(* CODESYS project Example9_PLC.project

Project tree, tasks and I/O mapping:
  Device : CODESYS Control Win V3, 3S - Smart Software Solutions GmbH, order no. 305021, version 3.5.7.0
    application Application
      libraries: Standard, * (System)
      task MainTask (cyclic, interval t#20ms, priority 1) calls PLC_PRG
      program PLC_PRG [ST]
      global variables GVL
      function block FB_G4LTL [ST]
    Ethernet : Ethernet, 3S - Smart Software Solutions GmbH, version 3.5.7.0
      Modbus_TCP_Master : Modbus TCP Master, 3S - Smart Software Solutions GmbH, version 3.5.6.0
          settings: AutoReconnect = TRUE
        Modbus_TCP_Slave : Modbus TCP Slave, 3S - Smart Software Solutions GmbH, version 3.5.7.0
            settings: Unit-ID = 1; IPAddress = [127, 0, 0, 1]; Channel 0.Function Code = 4; Channel 0.Read Offset = 16#0000; Channel 0.Read Length = 1; Channel 0.Write Offset = 0; Channel 0.Write Length = 0; Channel 0.Cycle Time = 100; Channel 1.Function Code = 4; Channel 1.Read Offset = 16#0001; Channel 1.Read Length = 1; Channel 1.Write Offset = 0; Channel 1.Write Length = 0; Channel 1.Cycle Time = 100; Channel 2.Function Code = 4; Channel 2.Read Offset = 16#0002; Channel 2.Read Length = 1; Channel 2.Write Offset = 0; Channel 2.Write Length = 0; Channel 2.Cycle Time = 100; Channel 3.Function Code = 4; Channel 3.Read Offset = 16#0003; Channel 3.Read Length = 1; Channel 3.Write Offset = 0; Channel 3.Write Length = 0; Channel 3.Cycle Time = 100; Channel 4.Function Code = 4; Channel 4.Read Offset = 16#0004; Channel 4.Read Length = 1; Channel 4.Write Offset = 0; Channel 4.Write Length = 0; Channel 4.Cycle Time = 100; Channel 5.Function Code = 6; Channel 5.Read Offset = 0; Channel 5.Read Length = 0; Channel 5.Write Offset = 16#0000; Channel 5.Write Length = 1; Channel 5.Cycle Time = 100; Channel 6.Function Code = 6; Channel 6.Read Offset = 0;
              Channel 6.Read Length = 0; Channel 6.Write Offset = 16#0002; Channel 6.Write Length = 1; Channel 6.Cycle Time = 100; Channel 7.Function Code = 6; Channel 7.Read Offset = 0; Channel 7.Read Length = 0; Channel 7.Write Offset = 16#0003; Channel 7.Write Length = 1; Channel 7.Cycle Time = 100; Channel 8.Function Code = 6; Channel 8.Read Offset = 0; Channel 8.Read Length = 0; Channel 8.Write Offset = 16#0004; Channel 8.Write Length = 1; Channel 8.Cycle Time = 100; Channel 9.Function Code = 6; Channel 9.Read Offset = 0; Channel 9.Read Length = 0; Channel 9.Write Offset = 16#0001; Channel 9.Write Length = 1; Channel 9.Cycle Time = 100
            input  Application.dIn0 : BOOL  // Channel 0.Channel 0.Bit0
            input  Application.dIn1 : BOOL  // Channel 1.Channel 1.Bit0
            input  Application.dIn2 : BOOL  // Channel 2.Channel 2.Bit0
            input  Application.dIn3 : BOOL  // Channel 3.Channel 3.Bit0
            input  Application.dIn4 : BOOL  // Channel 4.Channel 4.Bit0
            output Application.dOut0 : BOOL  // Channel 5.Channel 5.Bit0
            output Application.dOut2 : BOOL  // Channel 6.Channel 6.Bit0
            output Application.dOut3 : BOOL  // Channel 7.Channel 7.Bit0
            output Application.dOut4 : BOOL  // Channel 8.Channel 8.Bit0
            output Application.dOut1 : BOOL  // Channel 9.Channel 9.Bit0
            unmapped channels: Channel 0, Channel 1, Channel 2, Channel 3, Channel 4, Channel 5, Channel 6, Channel 7, Channel 8, Channel 9
*)

// Device/Application/GVL
VAR_GLOBAL
	
dIn0 : BOOL;
dIn1 : BOOL;
dIn2 : BOOL;
dIn3 : BOOL;
dIn4 : BOOL;

dOut0 : BOOL;
dOut1 : BOOL; 
dOut2 : BOOL; 
dOut3 : BOOL; 
dOut4 : BOOL; 
END_VAR

// Device/Application/PLC_PRG
PROGRAM PLC_PRG
VAR 
	fb: FB_G4LTL;	
END_VAR



// Direct looping
// Assign pins (from global variable to function block) 
fb.x0 := dIn0;

// Assign pins (from function block to global variable)
dOut0 := fb.y0;
dOut1 := fb.y1;
dOut2 := fb.y2;

// Run the function block
fb();

END_PROGRAM

// Device/Application/FB_G4LTL
FUNCTION_BLOCK FB_G4LTL
 (* Variable definition *)
   VAR_INPUT
      x0	: BOOL;
   END_VAR
   VAR_OUTPUT
      y0	: BOOL;
      y1	: BOOL;
      y2	: BOOL;
   END_VAR
   VAR
   (* The total number of states equals to 11 *)
      cstate16	: LINT := 0;
      t0	: TON;
      t0_reset	: BOOL := FALSE;
      t0_up	: BOOL := FALSE;
      t0_start	: BOOL := FALSE;
      t1	: TON;
      t1_reset	: BOOL := FALSE;
      t1_up	: BOOL := FALSE;
      t1_start	: BOOL := FALSE;	  
	  
	  T0_VALUE	: TIME := TIME#10S;
      T1_VALUE	: TIME := TIME#5s;
   END_VAR
   (* Constant definition  *)

CASE cstate16 OF
48641:
    IF ((x0 = FALSE) AND  (t0.Q = FALSE) AND  (t1.Q = FALSE)) THEN 
        cstate16 := 34931; y0 := FALSE; y1 := FALSE; y2 := FALSE; t0_start := FALSE;t1_start := FALSE; 
    ELSIF ((x0 = FALSE) AND  (t0.Q = FALSE) AND  (t1.Q = TRUE)) THEN 
        cstate16 := 34932; y0 := FALSE; y1 := FALSE; y2 := FALSE; t0_start := FALSE;t1_start := FALSE; 
    ELSIF ((x0 = FALSE) AND  (t0.Q = TRUE) AND  (t1.Q = FALSE)) THEN 
        cstate16 := 27731; y0 := FALSE; y1 := FALSE; y2 := FALSE; t0_start := FALSE;t1_start := TRUE; t1_up := FALSE; 
    ELSIF ((x0 = FALSE) AND  (t0.Q = TRUE) AND  (t1.Q = TRUE)) THEN 
        cstate16 := 27732; y0 := FALSE; y1 := FALSE; y2 := FALSE; t0_start := FALSE;t1_start := TRUE; t1_up := FALSE; 
    ELSIF ((x0 = TRUE) AND  (t0.Q = FALSE) AND  (t1.Q = FALSE)) THEN 
        cstate16 := 48641; y0 := TRUE; y1 := TRUE; y2 := FALSE; t0_start := FALSE;t1_start := FALSE; 
    ELSIF ((x0 = TRUE) AND  (t0.Q = FALSE) AND  (t1.Q = TRUE)) THEN 
        cstate16 := 48646; y0 := TRUE; y1 := TRUE; y2 := TRUE; t0_start := FALSE;t1_start := FALSE; 
    ELSIF ((x0 = TRUE) AND  (t0.Q = TRUE) AND  (t1.Q = FALSE)) THEN 
        cstate16 := 42449; y0 := TRUE; y1 := TRUE; y2 := FALSE; t0_start := FALSE;t1_start := TRUE; t1_up := FALSE; 
    ELSIF ((x0 = TRUE) AND  (t0.Q = TRUE) AND  (t1.Q = TRUE)) THEN 
        cstate16 := 42453; y0 := TRUE; y1 := TRUE; y2 := TRUE; t0_start := FALSE;t1_start := TRUE; t1_up := FALSE; 
    END_IF;
46659:
    IF ((x0 = FALSE) AND  (t0.Q = FALSE) AND  (t1.Q = FALSE)) THEN 
        cstate16 := 32883; y0 := FALSE; y1 := FALSE; y2 := FALSE; t0_start := FALSE;t1_start := FALSE; 
    ELSIF ((x0 = FALSE) AND  (t0.Q = FALSE) AND  (t1.Q = TRUE)) THEN 
        cstate16 := 34932; y0 := FALSE; y1 := FALSE; y2 := FALSE; t0_start := FALSE;t1_start := FALSE; 
    ELSIF ((x0 = FALSE) AND  (t0.Q = TRUE) AND  (t1.Q = FALSE)) THEN 
        cstate16 := 27763; y0 := FALSE; y1 := FALSE; y2 := FALSE; t0_start := FALSE;t1_start := FALSE; 
    ELSIF ((x0 = FALSE) AND  (t0.Q = TRUE) AND  (t1.Q = TRUE)) THEN 
        cstate16 := 28788; y0 := FALSE; y1 := FALSE; y2 := FALSE; t0_start := FALSE;t1_start := FALSE; 
    ELSIF ((x0 = TRUE) AND  (t0.Q = FALSE) AND  (t1.Q = FALSE)) THEN 
        cstate16 := 41187; y0 := TRUE; y1 := FALSE; y2 := FALSE; t0_start := TRUE; t0_up := FALSE;t1_start := FALSE; 
    ELSIF ((x0 = TRUE) AND  (t0.Q = FALSE) AND  (t1.Q = TRUE)) THEN 
        cstate16 := 40167; y0 := TRUE; y1 := FALSE; y2 := TRUE; t0_start := TRUE; t0_up := FALSE;t1_start := FALSE; 
    ELSIF ((x0 = TRUE) AND  (t0.Q = TRUE) AND  (t1.Q = FALSE)) THEN 
        cstate16 := 46659; y0 := TRUE; y1 := FALSE; y2 := FALSE; t0_start := FALSE;t1_start := FALSE; 
    ELSIF ((x0 = TRUE) AND  (t0.Q = TRUE) AND  (t1.Q = TRUE)) THEN 
        cstate16 := 47687; y0 := TRUE; y1 := FALSE; y2 := TRUE; t0_start := FALSE;t1_start := FALSE; 
    END_IF;
46651:
    IF ((x0 = FALSE) AND  (t0.Q = FALSE) AND  (t1.Q = FALSE)) THEN 
        cstate16 := 32883; y0 := FALSE; y1 := FALSE; y2 := FALSE; t0_start := FALSE;t1_start := FALSE; 
    ELSIF ((x0 = FALSE) AND  (t0.Q = FALSE) AND  (t1.Q = TRUE)) THEN 
        cstate16 := 34932; y0 := FALSE; y1 := FALSE; y2 := FALSE; t0_start := FALSE;t1_start := FALSE; 
    ELSIF ((x0 = FALSE) AND  (t0.Q = TRUE) AND  (t1.Q = FALSE)) THEN 
        cstate16 := 27763; y0 := FALSE; y1 := FALSE; y2 := FALSE; t0_start := FALSE;t1_start := FALSE; 
    ELSIF ((x0 = FALSE) AND  (t0.Q = TRUE) AND  (t1.Q = TRUE)) THEN 
        cstate16 := 28788; y0 := FALSE; y1 := FALSE; y2 := FALSE; t0_start := FALSE;t1_start := FALSE; 
    ELSIF ((x0 = TRUE) AND  (t0.Q = FALSE) AND  (t1.Q = FALSE)) THEN 
        cstate16 := 41643; y0 := TRUE; y1 := TRUE; y2 := TRUE; t0_start := TRUE; t0_up := FALSE;t1_start := FALSE; 
    ELSIF ((x0 = TRUE) AND  (t0.Q = FALSE) AND  (t1.Q = TRUE)) THEN 
        cstate16 := 40647; y0 := TRUE; y1 := TRUE; y2 := TRUE; t0_start := TRUE; t0_up := FALSE;t1_start := FALSE; 
    ELSIF ((x0 = TRUE) AND  (t0.Q = TRUE) AND  (t1.Q = FALSE)) THEN 
        cstate16 := 46747; y0 := TRUE; y1 := TRUE; y2 := TRUE; t0_start := FALSE;t1_start := FALSE; 
    ELSIF ((x0 = TRUE) AND  (t0.Q = TRUE) AND  (t1.Q = TRUE)) THEN 
        cstate16 := 47799; y0 := TRUE; y1 := TRUE; y2 := TRUE; t0_start := FALSE;t1_start := FALSE; 
    END_IF;
25798:
    IF ((x0 = FALSE) AND  (t0.Q = FALSE) AND  (t1.Q = FALSE)) THEN 
        cstate16 := 26739; y0 := FALSE; y1 := FALSE; y2 := FALSE; t0_start := FALSE;t1_start := FALSE; 
    ELSIF ((x0 = FALSE) AND  (t0.Q = FALSE) AND  (t1.Q = TRUE)) THEN 
        cstate16 := 26740; y0 := FALSE; y1 := FALSE; y2 := FALSE; t0_start := FALSE;t1_start := FALSE; 
    ELSIF ((x0 = FALSE) AND  (t0.Q = TRUE) AND  (t1.Q = FALSE)) THEN 
        cstate16 := 17491; y0 := FALSE; y1 := FALSE; y2 := FALSE; t0_start := FALSE;t1_start := TRUE; t1_up := FALSE; 
    ELSIF ((x0 = FALSE) AND  (t0.Q = TRUE) AND  (t1.Q = TRUE)) THEN 
        cstate16 := 17492; y0 := FALSE; y1 := FALSE; y2 := FALSE; t0_start := FALSE;t1_start := TRUE; t1_up := FALSE; 
    ELSIF ((x0 = TRUE) AND  (t0.Q = FALSE) AND  (t1.Q = FALSE)) THEN 
        cstate16 := 26042; y0 := TRUE; y1 := FALSE; y2 := TRUE; t0_start := FALSE;t1_start := FALSE; 
    ELSIF ((x0 = TRUE) AND  (t0.Q = FALSE) AND  (t1.Q = TRUE)) THEN 
        cstate16 := 26038; y0 := TRUE; y1 := FALSE; y2 := TRUE; t0_start := FALSE;t1_start := FALSE; 
    ELSIF ((x0 = TRUE) AND  (t0.Q = TRUE) AND  (t1.Q = FALSE)) THEN 
        cstate16 := 42457; y0 := TRUE; y1 := TRUE; y2 := TRUE; t0_start := FALSE;t1_start := TRUE; t1_up := FALSE; 
    ELSIF ((x0 = TRUE) AND  (t0.Q = TRUE) AND  (t1.Q = TRUE)) THEN 
        cstate16 := 42453; y0 := TRUE; y1 := TRUE; y2 := TRUE; t0_start := FALSE;t1_start := TRUE; t1_up := FALSE; 
    END_IF;
34931:
    IF ((x0 = FALSE) AND  (t0.Q = FALSE) AND  (t1.Q = FALSE)) THEN 
        cstate16 := 34931; y0 := FALSE; y1 := FALSE; y2 := FALSE; t0_start := FALSE;t1_start := FALSE; 
    ELSIF ((x0 = FALSE) AND  (t0.Q = FALSE) AND  (t1.Q = TRUE)) THEN 
        cstate16 := 34932; y0 := FALSE; y1 := FALSE; y2 := FALSE; t0_start := FALSE;t1_start := FALSE; 
    ELSIF ((x0 = FALSE) AND  (t0.Q = TRUE) AND  (t1.Q = FALSE)) THEN 
        cstate16 := 27731; y0 := FALSE; y1 := FALSE; y2 := FALSE; t0_start := FALSE;t1_start := TRUE; t1_up := FALSE; 
    ELSIF ((x0 = FALSE) AND  (t0.Q = TRUE) AND  (t1.Q = TRUE)) THEN 
        cstate16 := 27732; y0 := FALSE; y1 := FALSE; y2 := FALSE; t0_start := FALSE;t1_start := TRUE; t1_up := FALSE; 
    ELSIF ((x0 = TRUE) AND  (t0.Q = FALSE) AND  (t1.Q = FALSE)) THEN 
        cstate16 := 40163; y0 := TRUE; y1 := FALSE; y2 := FALSE; t0_start := TRUE; t0_up := FALSE;t1_start := FALSE; 
    ELSIF ((x0 = TRUE) AND  (t0.Q = FALSE) AND  (t1.Q = TRUE)) THEN 
        cstate16 := 40167; y0 := TRUE; y1 := FALSE; y2 := TRUE; t0_start := TRUE; t0_up := FALSE;t1_start := FALSE; 
    ELSIF ((x0 = TRUE) AND  (t0.Q = TRUE) AND  (t1.Q = FALSE)) THEN 
        cstate16 := 38147; y0 := TRUE; y1 := TRUE; y2 := FALSE; t0_start := TRUE; t0_up := FALSE;t1_start := TRUE; t1_up := FALSE; 
    ELSIF ((x0 = TRUE) AND  (t0.Q = TRUE) AND  (t1.Q = TRUE)) THEN 
        cstate16 := 38152; y0 := TRUE; y1 := TRUE; y2 := TRUE; t0_start := TRUE; t0_up := FALSE;t1_start := TRUE; t1_up := FALSE; 
    END_IF;
47687:
    IF ((x0 = FALSE) AND  (t0.Q = FALSE) AND  (t1.Q = FALSE)) THEN 
        cstate16 := 34931; y0 := FALSE; y1 := FALSE; y2 := FALSE; t0_start := FALSE;t1_start := FALSE; 
    ELSIF ((x0 = FALSE) AND  (t0.Q = FALSE) AND  (t1.Q = TRUE)) THEN 
        cstate16 := 34932; y0 := FALSE; y1 := FALSE; y2 := FALSE; t0_start := FALSE;t1_start := FALSE; 
    ELSIF ((x0 = FALSE) AND  (t0.Q = TRUE) AND  (t1.Q = FALSE)) THEN 
        cstate16 := 28787; y0 := FALSE; y1 := FALSE; y2 := FALSE; t0_start := FALSE;t1_start := FALSE; 
    ELSIF ((x0 = FALSE) AND  (t0.Q = TRUE) AND  (t1.Q = TRUE)) THEN 
        cstate16 := 28788; y0 := FALSE; y1 := FALSE; y2 := FALSE; t0_start := FALSE;t1_start := FALSE; 
    ELSIF ((x0 = TRUE) AND  (t0.Q = FALSE) AND  (t1.Q = FALSE)) THEN 
        cstate16 := 40172; y0 := TRUE; y1 := FALSE; y2 := TRUE; t0_start := TRUE; t0_up := FALSE;t1_start := FALSE; 
    ELSIF ((x0 = TRUE) AND  (t0.Q = FALSE) AND  (t1.Q = TRUE)) THEN 
        cstate16 := 40167; y0 := TRUE; y1 := FALSE; y2 := TRUE; t0_start := TRUE; t0_up := FALSE;t1_start := FALSE; 
    ELSIF ((x0 = TRUE) AND  (t0.Q = TRUE) AND  (t1.Q = FALSE)) THEN 
        cstate16 := 47692; y0 := TRUE; y1 := FALSE; y2 := TRUE; t0_start := FALSE;t1_start := FALSE; 
    ELSIF ((x0 = TRUE) AND  (t0.Q = TRUE) AND  (t1.Q = TRUE)) THEN 
        cstate16 := 47687; y0 := TRUE; y1 := FALSE; y2 := TRUE; t0_start := FALSE;t1_start := FALSE; 
    END_IF;
43409:
    IF ((x0 = FALSE) AND  (t0.Q = FALSE) AND  (t1.Q = FALSE)) THEN 
        cstate16 := 34931; y0 := FALSE; y1 := FALSE; y2 := FALSE; t0_start := FALSE;t1_start := FALSE; 
    ELSIF ((x0 = FALSE) AND  (t0.Q = FALSE) AND  (t1.Q = TRUE)) THEN 
        cstate16 := 34932; y0 := FALSE; y1 := FALSE; y2 := FALSE; t0_start := FALSE;t1_start := FALSE; 
    ELSIF ((x0 = FALSE) AND  (t0.Q = TRUE) AND  (t1.Q = FALSE)) THEN 
        cstate16 := 28787; y0 := FALSE; y1 := FALSE; y2 := FALSE; t0_start := FALSE;t1_start := FALSE; 
    ELSIF ((x0 = FALSE) AND  (t0.Q = TRUE) AND  (t1.Q = TRUE)) THEN 
        cstate16 := 28788; y0 := FALSE; y1 := FALSE; y2 := FALSE; t0_start := FALSE;t1_start := FALSE; 
    ELSIF ((x0 = TRUE) AND  (t0.Q = FALSE) AND  (t1.Q = FALSE)) THEN 
        cstate16 := 48529; y0 := TRUE; y1 := FALSE; y2 := FALSE; t0_start := FALSE;t1_start := FALSE; 
    ELSIF ((x0 = TRUE) AND  (t0.Q = FALSE) AND  (t1.Q = TRUE)) THEN 
        cstate16 := 48534; y0 := TRUE; y1 := FALSE; y2 := TRUE; t0_start := FALSE;t1_start := FALSE; 
    ELSIF ((x0 = TRUE) AND  (t0.Q = TRUE) AND  (t1.Q = FALSE)) THEN 
        cstate16 := 43409; y0 := TRUE; y1 := FALSE; y2 := FALSE; t0_start := FALSE;t1_start := FALSE; 
    ELSIF ((x0 = TRUE) AND  (t0.Q = TRUE) AND  (t1.Q = TRUE)) THEN 
        cstate16 := 43414; y0 := TRUE; y1 := FALSE; y2 := TRUE; t0_start := FALSE;t1_start := FALSE; 
    END_IF;
34932:
    IF ((x0 = FALSE) AND  (t0.Q = FALSE) AND  (t1.Q = FALSE)) THEN 
        cstate16 := 34931; y0 := FALSE; y1 := FALSE; y2 := FALSE; t0_start := FALSE;t1_start := FALSE; 
    ELSIF ((x0 = FALSE) AND  (t0.Q = FALSE) AND  (t1.Q = TRUE)) THEN 
        cstate16 := 34932; y0 := FALSE; y1 := FALSE; y2 := FALSE; t0_start := FALSE;t1_start := FALSE; 
    ELSIF ((x0 = FALSE) AND  (t0.Q = TRUE) AND  (t1.Q = FALSE)) THEN 
        cstate16 := 27731; y0 := FALSE; y1 := FALSE; y2 := FALSE; t0_start := FALSE;t1_start := TRUE; t1_up := FALSE; 
    ELSIF ((x0 = FALSE) AND  (t0.Q = TRUE) AND  (t1.Q = TRUE)) THEN 
        cstate16 := 27732; y0 := FALSE; y1 := FALSE; y2 := FALSE; t0_start := FALSE;t1_start := TRUE; t1_up := FALSE; 
    ELSIF ((x0 = TRUE) AND  (t0.Q = FALSE) AND  (t1.Q = FALSE)) THEN 
        cstate16 := 40163; y0 := TRUE; y1 := FALSE; y2 := FALSE; t0_start := TRUE; t0_up := FALSE;t1_start := FALSE; 
    ELSIF ((x0 = TRUE) AND  (t0.Q = FALSE) AND  (t1.Q = TRUE)) THEN 
        cstate16 := 40164; y0 := TRUE; y1 := FALSE; y2 := FALSE; t0_start := TRUE; t0_up := FALSE;t1_start := FALSE; 
    ELSIF ((x0 = TRUE) AND  (t0.Q = TRUE) AND  (t1.Q = FALSE)) THEN 
        cstate16 := 38147; y0 := TRUE; y1 := TRUE; y2 := FALSE; t0_start := TRUE; t0_up := FALSE;t1_start := TRUE; t1_up := FALSE; 
    ELSIF ((x0 = TRUE) AND  (t0.Q = TRUE) AND  (t1.Q = TRUE)) THEN 
        cstate16 := 38148; y0 := TRUE; y1 := TRUE; y2 := FALSE; t0_start := TRUE; t0_up := FALSE;t1_start := TRUE; t1_up := FALSE; 
    END_IF;
6209:
    IF ((x0 = FALSE) AND  (t0.Q = FALSE) AND  (t1.Q = FALSE)) THEN 
        cstate16 := 34931; y0 := FALSE; y1 := FALSE; y2 := FALSE; t0_start := FALSE;t1_start := FALSE; 
    ELSIF ((x0 = FALSE) AND  (t0.Q = FALSE) AND  (t1.Q = TRUE)) THEN 
        cstate16 := 34932; y0 := FALSE; y1 := FALSE; y2 := FALSE; t0_start := FALSE;t1_start := FALSE; 
    ELSIF ((x0 = FALSE) AND  (t0.Q = TRUE) AND  (t1.Q = FALSE)) THEN 
        cstate16 := 28787; y0 := FALSE; y1 := FALSE; y2 := FALSE; t0_start := FALSE;t1_start := FALSE; 
    ELSIF ((x0 = FALSE) AND  (t0.Q = TRUE) AND  (t1.Q = TRUE)) THEN 
        cstate16 := 28788; y0 := FALSE; y1 := FALSE; y2 := FALSE; t0_start := FALSE;t1_start := FALSE; 
    ELSIF ((x0 = TRUE) AND  (t0.Q = FALSE) AND  (t1.Q = FALSE)) THEN 
        cstate16 := 14401; y0 := FALSE; y1 := FALSE; y2 := FALSE; t0_start := FALSE;t1_start := FALSE; 
    ELSIF ((x0 = TRUE) AND  (t0.Q = FALSE) AND  (t1.Q = TRUE)) THEN 
        cstate16 := 14406; y0 := FALSE; y1 := FALSE; y2 := TRUE; t0_start := FALSE;t1_start := FALSE; 
    ELSIF ((x0 = TRUE) AND  (t0.Q = TRUE) AND  (t1.Q = FALSE)) THEN 
        cstate16 := 6209; y0 := FALSE; y1 := FALSE; y2 := FALSE; t0_start := FALSE;t1_start := FALSE; 
    ELSIF ((x0 = TRUE) AND  (t0.Q = TRUE) AND  (t1.Q = TRUE)) THEN 
        cstate16 := 6214; y0 := FALSE; y1 := FALSE; y2 := TRUE; t0_start := FALSE;t1_start := FALSE; 
    END_IF;
42489:
    IF ((x0 = FALSE) AND  (t0.Q = FALSE) AND  (t1.Q = FALSE)) THEN 
        cstate16 := 32883; y0 := FALSE; y1 := FALSE; y2 := FALSE; t0_start := FALSE;t1_start := FALSE; 
    ELSIF ((x0 = FALSE) AND  (t0.Q = FALSE) AND  (t1.Q = TRUE)) THEN 
        cstate16 := 34932; y0 := FALSE; y1 := FALSE; y2 := FALSE; t0_start := FALSE;t1_start := FALSE; 
    ELSIF ((x0 = FALSE) AND  (t0.Q = TRUE) AND  (t1.Q = FALSE)) THEN 
        cstate16 := 27763; y0 := FALSE; y1 := FALSE; y2 := FALSE; t0_start := FALSE;t1_start := FALSE; 
    ELSIF ((x0 = FALSE) AND  (t0.Q = TRUE) AND  (t1.Q = TRUE)) THEN 
        cstate16 := 28788; y0 := FALSE; y1 := FALSE; y2 := FALSE; t0_start := FALSE;t1_start := FALSE; 
    ELSIF ((x0 = TRUE) AND  (t0.Q = FALSE) AND  (t1.Q = FALSE)) THEN 
        cstate16 := 49657; y0 := TRUE; y1 := TRUE; y2 := TRUE; t0_start := FALSE;t1_start := FALSE; 
    ELSIF ((x0 = TRUE) AND  (t0.Q = FALSE) AND  (t1.Q = TRUE)) THEN 
        cstate16 := 48646; y0 := TRUE; y1 := TRUE; y2 := TRUE; t0_start := FALSE;t1_start := FALSE; 
    ELSIF ((x0 = TRUE) AND  (t0.Q = TRUE) AND  (t1.Q = FALSE)) THEN 
        cstate16 := 42489; y0 := TRUE; y1 := TRUE; y2 := TRUE; t0_start := FALSE;t1_start := FALSE; 
    ELSIF ((x0 = TRUE) AND  (t0.Q = TRUE) AND  (t1.Q = TRUE)) THEN 
        cstate16 := 43526; y0 := TRUE; y1 := TRUE; y2 := TRUE; t0_start := FALSE;t1_start := FALSE; 
    END_IF;
6490:
    IF ((x0 = FALSE) AND  (t0.Q = FALSE) AND  (t1.Q = FALSE)) THEN 
        cstate16 := 34931; y0 := FALSE; y1 := FALSE; y2 := FALSE; t0_start := FALSE;t1_start := FALSE; 
    ELSIF ((x0 = FALSE) AND  (t0.Q = FALSE) AND  (t1.Q = TRUE)) THEN 
        cstate16 := 34932; y0 := FALSE; y1 := FALSE; y2 := FALSE; t0_start := FALSE;t1_start := FALSE; 
    ELSIF ((x0 = FALSE) AND  (t0.Q = TRUE) AND  (t1.Q = FALSE)) THEN 
        cstate16 := 28787; y0 := FALSE; y1 := FALSE; y2 := FALSE; t0_start := FALSE;t1_start := FALSE; 
    ELSIF ((x0 = FALSE) AND  (t0.Q = TRUE) AND  (t1.Q = TRUE)) THEN 
        cstate16 := 28788; y0 := FALSE; y1 := FALSE; y2 := FALSE; t0_start := FALSE;t1_start := FALSE; 
    ELSIF ((x0 = TRUE) AND  (t0.Q = FALSE) AND  (t1.Q = FALSE)) THEN 
        cstate16 := 14682; y0 := FALSE; y1 := TRUE; y2 := TRUE; t0_start := FALSE;t1_start := FALSE; 
    ELSIF ((x0 = TRUE) AND  (t0.Q = FALSE) AND  (t1.Q = TRUE)) THEN 
        cstate16 := 14678; y0 := FALSE; y1 := TRUE; y2 := TRUE; t0_start := FALSE;t1_start := FALSE; 
    ELSIF ((x0 = TRUE) AND  (t0.Q = TRUE) AND  (t1.Q = FALSE)) THEN 
        cstate16 := 6490; y0 := FALSE; y1 := TRUE; y2 := TRUE; t0_start := FALSE;t1_start := FALSE; 
    ELSIF ((x0 = TRUE) AND  (t0.Q = TRUE) AND  (t1.Q = TRUE)) THEN 
        cstate16 := 6486; y0 := FALSE; y1 := TRUE; y2 := TRUE; t0_start := FALSE;t1_start := FALSE; 
    END_IF;
6210:
    IF ((x0 = FALSE) AND  (t0.Q = FALSE) AND  (t1.Q = FALSE)) THEN 
        cstate16 := 34931; y0 := FALSE; y1 := FALSE; y2 := FALSE; t0_start := FALSE;t1_start := FALSE; 
    ELSIF ((x0 = FALSE) AND  (t0.Q = FALSE) AND  (t1.Q = TRUE)) THEN 
        cstate16 := 34932; y0 := FALSE; y1 := FALSE; y2 := FALSE; t0_start := FALSE;t1_start := FALSE; 
    ELSIF ((x0 = FALSE) AND  (t0.Q = TRUE) AND  (t1.Q = FALSE)) THEN 
        cstate16 := 28787; y0 := FALSE; y1 := FALSE; y2 := FALSE; t0_start := FALSE;t1_start := FALSE; 
    ELSIF ((x0 = FALSE) AND  (t0.Q = TRUE) AND  (t1.Q = TRUE)) THEN 
        cstate16 := 28788; y0 := FALSE; y1 := FALSE; y2 := FALSE; t0_start := FALSE;t1_start := FALSE; 
    ELSIF ((x0 = TRUE) AND  (t0.Q = FALSE) AND  (t1.Q = FALSE)) THEN 
        cstate16 := 14401; y0 := FALSE; y1 := FALSE; y2 := FALSE; t0_start := FALSE;t1_start := FALSE; 
    ELSIF ((x0 = TRUE) AND  (t0.Q = FALSE) AND  (t1.Q = TRUE)) THEN 
        cstate16 := 14402; y0 := FALSE; y1 := FALSE; y2 := FALSE; t0_start := FALSE;t1_start := FALSE; 
    ELSIF ((x0 = TRUE) AND  (t0.Q = TRUE) AND  (t1.Q = FALSE)) THEN 
        cstate16 := 6209; y0 := FALSE; y1 := FALSE; y2 := FALSE; t0_start := FALSE;t1_start := FALSE; 
    ELSIF ((x0 = TRUE) AND  (t0.Q = TRUE) AND  (t1.Q = TRUE)) THEN 
        cstate16 := 6210; y0 := FALSE; y1 := FALSE; y2 := FALSE; t0_start := FALSE;t1_start := FALSE; 
    END_IF;
25794:
    IF ((x0 = FALSE) AND  (t0.Q = FALSE) AND  (t1.Q = FALSE)) THEN 
        cstate16 := 26739; y0 := FALSE; y1 := FALSE; y2 := FALSE; t0_start := FALSE;t1_start := FALSE; 
    ELSIF ((x0 = FALSE) AND  (t0.Q = FALSE) AND  (t1.Q = TRUE)) THEN 
        cstate16 := 26740; y0 := FALSE; y1 := FALSE; y2 := FALSE; t0_start := FALSE;t1_start := FALSE; 
    ELSIF ((x0 = FALSE) AND  (t0.Q = TRUE) AND  (t1.Q = FALSE)) THEN 
        cstate16 := 17491; y0 := FALSE; y1 := FALSE; y2 := FALSE; t0_start := FALSE;t1_start := TRUE; t1_up := FALSE; 
    ELSIF ((x0 = FALSE) AND  (t0.Q = TRUE) AND  (t1.Q = TRUE)) THEN 
        cstate16 := 17492; y0 := FALSE; y1 := FALSE; y2 := FALSE; t0_start := FALSE;t1_start := TRUE; t1_up := FALSE; 
    ELSIF ((x0 = TRUE) AND  (t0.Q = FALSE) AND  (t1.Q = FALSE)) THEN 
        cstate16 := 26033; y0 := TRUE; y1 := FALSE; y2 := FALSE; t0_start := FALSE;t1_start := FALSE; 
    ELSIF ((x0 = TRUE) AND  (t0.Q = FALSE) AND  (t1.Q = TRUE)) THEN 
        cstate16 := 26034; y0 := TRUE; y1 := FALSE; y2 := FALSE; t0_start := FALSE;t1_start := FALSE; 
    ELSIF ((x0 = TRUE) AND  (t0.Q = TRUE) AND  (t1.Q = FALSE)) THEN 
        cstate16 := 42449; y0 := TRUE; y1 := TRUE; y2 := FALSE; t0_start := FALSE;t1_start := TRUE; t1_up := FALSE; 
    ELSIF ((x0 = TRUE) AND  (t0.Q = TRUE) AND  (t1.Q = TRUE)) THEN 
        cstate16 := 42450; y0 := TRUE; y1 := TRUE; y2 := FALSE; t0_start := FALSE;t1_start := TRUE; t1_up := FALSE; 
    END_IF;
25793:
    IF ((x0 = FALSE) AND  (t0.Q = FALSE) AND  (t1.Q = FALSE)) THEN 
        cstate16 := 26739; y0 := FALSE; y1 := FALSE; y2 := FALSE; t0_start := FALSE;t1_start := FALSE; 
    ELSIF ((x0 = FALSE) AND  (t0.Q = FALSE) AND  (t1.Q = TRUE)) THEN 
        cstate16 := 26740; y0 := FALSE; y1 := FALSE; y2 := FALSE; t0_start := FALSE;t1_start := FALSE; 
    ELSIF ((x0 = FALSE) AND  (t0.Q = TRUE) AND  (t1.Q = FALSE)) THEN 
        cstate16 := 17491; y0 := FALSE; y1 := FALSE; y2 := FALSE; t0_start := FALSE;t1_start := TRUE; t1_up := FALSE; 
    ELSIF ((x0 = FALSE) AND  (t0.Q = TRUE) AND  (t1.Q = TRUE)) THEN 
        cstate16 := 17492; y0 := FALSE; y1 := FALSE; y2 := FALSE; t0_start := FALSE;t1_start := TRUE; t1_up := FALSE; 
    ELSIF ((x0 = TRUE) AND  (t0.Q = FALSE) AND  (t1.Q = FALSE)) THEN 
        cstate16 := 26033; y0 := TRUE; y1 := FALSE; y2 := FALSE; t0_start := FALSE;t1_start := FALSE; 
    ELSIF ((x0 = TRUE) AND  (t0.Q = FALSE) AND  (t1.Q = TRUE)) THEN 
        cstate16 := 26038; y0 := TRUE; y1 := FALSE; y2 := TRUE; t0_start := FALSE;t1_start := FALSE; 
    ELSIF ((x0 = TRUE) AND  (t0.Q = TRUE) AND  (t1.Q = FALSE)) THEN 
        cstate16 := 42449; y0 := TRUE; y1 := TRUE; y2 := FALSE; t0_start := FALSE;t1_start := TRUE; t1_up := FALSE; 
    ELSIF ((x0 = TRUE) AND  (t0.Q = TRUE) AND  (t1.Q = TRUE)) THEN 
        cstate16 := 42453; y0 := TRUE; y1 := TRUE; y2 := TRUE; t0_start := FALSE;t1_start := TRUE; t1_up := FALSE; 
    END_IF;
47683:
    IF ((x0 = FALSE) AND  (t0.Q = FALSE) AND  (t1.Q = FALSE)) THEN 
        cstate16 := 34931; y0 := FALSE; y1 := FALSE; y2 := FALSE; t0_start := FALSE;t1_start := FALSE; 
    ELSIF ((x0 = FALSE) AND  (t0.Q = FALSE) AND  (t1.Q = TRUE)) THEN 
        cstate16 := 34932; y0 := FALSE; y1 := FALSE; y2 := FALSE; t0_start := FALSE;t1_start := FALSE; 
    ELSIF ((x0 = FALSE) AND  (t0.Q = TRUE) AND  (t1.Q = FALSE)) THEN 
        cstate16 := 28787; y0 := FALSE; y1 := FALSE; y2 := FALSE; t0_start := FALSE;t1_start := FALSE; 
    ELSIF ((x0 = FALSE) AND  (t0.Q = TRUE) AND  (t1.Q = TRUE)) THEN 
        cstate16 := 28788; y0 := FALSE; y1 := FALSE; y2 := FALSE; t0_start := FALSE;t1_start := FALSE; 
    ELSIF ((x0 = TRUE) AND  (t0.Q = FALSE) AND  (t1.Q = FALSE)) THEN 
        cstate16 := 40163; y0 := TRUE; y1 := FALSE; y2 := FALSE; t0_start := TRUE; t0_up := FALSE;t1_start := FALSE; 
    ELSIF ((x0 = TRUE) AND  (t0.Q = FALSE) AND  (t1.Q = TRUE)) THEN 
        cstate16 := 40167; y0 := TRUE; y1 := FALSE; y2 := TRUE; t0_start := TRUE; t0_up := FALSE;t1_start := FALSE; 
    ELSIF ((x0 = TRUE) AND  (t0.Q = TRUE) AND  (t1.Q = FALSE)) THEN 
        cstate16 := 47683; y0 := TRUE; y1 := FALSE; y2 := FALSE; t0_start := FALSE;t1_start := FALSE; 
    ELSIF ((x0 = TRUE) AND  (t0.Q = TRUE) AND  (t1.Q = TRUE)) THEN 
        cstate16 := 47687; y0 := TRUE; y1 := FALSE; y2 := TRUE; t0_start := FALSE;t1_start := FALSE; 
    END_IF;
6214:
    IF ((x0 = FALSE) AND  (t0.Q = FALSE) AND  (t1.Q = FALSE)) THEN 
        cstate16 := 34931; y0 := FALSE; y1 := FALSE; y2 := FALSE; t0_start := FALSE;t1_start := FALSE; 
    ELSIF ((x0 = FALSE) AND  (t0.Q = FALSE) AND  (t1.Q = TRUE)) THEN 
        cstate16 := 34932; y0 := FALSE; y1 := FALSE; y2 := FALSE; t0_start := FALSE;t1_start := FALSE; 
    ELSIF ((x0 = FALSE) AND  (t0.Q = TRUE) AND  (t1.Q = FALSE)) THEN 
        cstate16 := 28787; y0 := FALSE; y1 := FALSE; y2 := FALSE; t0_start := FALSE;t1_start := FALSE; 
    ELSIF ((x0 = FALSE) AND  (t0.Q = TRUE) AND  (t1.Q = TRUE)) THEN 
        cstate16 := 28788; y0 := FALSE; y1 := FALSE; y2 := FALSE; t0_start := FALSE;t1_start := FALSE; 
    ELSIF ((x0 = TRUE) AND  (t0.Q = FALSE) AND  (t1.Q = FALSE)) THEN 
        cstate16 := 14410; y0 := FALSE; y1 := FALSE; y2 := TRUE; t0_start := FALSE;t1_start := FALSE; 
    ELSIF ((x0 = TRUE) AND  (t0.Q = FALSE) AND  (t1.Q = TRUE)) THEN 
        cstate16 := 14406; y0 := FALSE; y1 := FALSE; y2 := TRUE; t0_start := FALSE;t1_start := FALSE; 
    ELSIF ((x0 = TRUE) AND  (t0.Q = TRUE) AND  (t1.Q = FALSE)) THEN 
        cstate16 := 6218; y0 := FALSE; y1 := FALSE; y2 := TRUE; t0_start := FALSE;t1_start := FALSE; 
    ELSIF ((x0 = TRUE) AND  (t0.Q = TRUE) AND  (t1.Q = TRUE)) THEN 
        cstate16 := 6214; y0 := FALSE; y1 := FALSE; y2 := TRUE; t0_start := FALSE;t1_start := FALSE; 
    END_IF;
47684:
    IF ((x0 = FALSE) AND  (t0.Q = FALSE) AND  (t1.Q = FALSE)) THEN 
        cstate16 := 34931; y0 := FALSE; y1 := FALSE; y2 := FALSE; t0_start := FALSE;t1_start := FALSE; 
    ELSIF ((x0 = FALSE) AND  (t0.Q = FALSE) AND  (t1.Q = TRUE)) THEN 
        cstate16 := 34932; y0 := FALSE; y1 := FALSE; y2 := FALSE; t0_start := FALSE;t1_start := FALSE; 
    ELSIF ((x0 = FALSE) AND  (t0.Q = TRUE) AND  (t1.Q = FALSE)) THEN 
        cstate16 := 28787; y0 := FALSE; y1 := FALSE; y2 := FALSE; t0_start := FALSE;t1_start := FALSE; 
    ELSIF ((x0 = FALSE) AND  (t0.Q = TRUE) AND  (t1.Q = TRUE)) THEN 
        cstate16 := 28788; y0 := FALSE; y1 := FALSE; y2 := FALSE; t0_start := FALSE;t1_start := FALSE; 
    ELSIF ((x0 = TRUE) AND  (t0.Q = FALSE) AND  (t1.Q = FALSE)) THEN 
        cstate16 := 40163; y0 := TRUE; y1 := FALSE; y2 := FALSE; t0_start := TRUE; t0_up := FALSE;t1_start := FALSE; 
    ELSIF ((x0 = TRUE) AND  (t0.Q = FALSE) AND  (t1.Q = TRUE)) THEN 
        cstate16 := 40164; y0 := TRUE; y1 := FALSE; y2 := FALSE; t0_start := TRUE; t0_up := FALSE;t1_start := FALSE; 
    ELSIF ((x0 = TRUE) AND  (t0.Q = TRUE) AND  (t1.Q = FALSE)) THEN 
        cstate16 := 47683; y0 := TRUE; y1 := FALSE; y2 := FALSE; t0_start := FALSE;t1_start := FALSE; 
    ELSIF ((x0 = TRUE) AND  (t0.Q = TRUE) AND  (t1.Q = TRUE)) THEN 
        cstate16 := 47684; y0 := TRUE; y1 := FALSE; y2 := FALSE; t0_start := FALSE;t1_start := FALSE; 
    END_IF;
42481:
    IF ((x0 = FALSE) AND  (t0.Q = FALSE) AND  (t1.Q = FALSE)) THEN 
        cstate16 := 32883; y0 := FALSE; y1 := FALSE; y2 := FALSE; t0_start := FALSE;t1_start := FALSE; 
    ELSIF ((x0 = FALSE) AND  (t0.Q = FALSE) AND  (t1.Q = TRUE)) THEN 
        cstate16 := 34932; y0 := FALSE; y1 := FALSE; y2 := FALSE; t0_start := FALSE;t1_start := FALSE; 
    ELSIF ((x0 = FALSE) AND  (t0.Q = TRUE) AND  (t1.Q = FALSE)) THEN 
        cstate16 := 27763; y0 := FALSE; y1 := FALSE; y2 := FALSE; t0_start := FALSE;t1_start := FALSE; 
    ELSIF ((x0 = FALSE) AND  (t0.Q = TRUE) AND  (t1.Q = TRUE)) THEN 
        cstate16 := 28788; y0 := FALSE; y1 := FALSE; y2 := FALSE; t0_start := FALSE;t1_start := FALSE; 
    ELSIF ((x0 = TRUE) AND  (t0.Q = FALSE) AND  (t1.Q = FALSE)) THEN 
        cstate16 := 49649; y0 := TRUE; y1 := TRUE; y2 := FALSE; t0_start := FALSE;t1_start := FALSE; 
    ELSIF ((x0 = TRUE) AND  (t0.Q = FALSE) AND  (t1.Q = TRUE)) THEN 
        cstate16 := 48646; y0 := TRUE; y1 := TRUE; y2 := TRUE; t0_start := FALSE;t1_start := FALSE; 
    ELSIF ((x0 = TRUE) AND  (t0.Q = TRUE) AND  (t1.Q = FALSE)) THEN 
        cstate16 := 42481; y0 := TRUE; y1 := TRUE; y2 := FALSE; t0_start := FALSE;t1_start := FALSE; 
    ELSIF ((x0 = TRUE) AND  (t0.Q = TRUE) AND  (t1.Q = TRUE)) THEN 
        cstate16 := 43526; y0 := TRUE; y1 := TRUE; y2 := TRUE; t0_start := FALSE;t1_start := FALSE; 
    END_IF;
48646:
    IF ((x0 = FALSE) AND  (t0.Q = FALSE) AND  (t1.Q = FALSE)) THEN 
        cstate16 := 34931; y0 := FALSE; y1 := FALSE; y2 := FALSE; t0_start := FALSE;t1_start := FALSE; 
    ELSIF ((x0 = FALSE) AND  (t0.Q = FALSE) AND  (t1.Q = TRUE)) THEN 
        cstate16 := 34932; y0 := FALSE; y1 := FALSE; y2 := FALSE; t0_start := FALSE;t1_start := FALSE; 
    ELSIF ((x0 = FALSE) AND  (t0.Q = TRUE) AND  (t1.Q = FALSE)) THEN 
        cstate16 := 27731; y0 := FALSE; y1 := FALSE; y2 := FALSE; t0_start := FALSE;t1_start := TRUE; t1_up := FALSE; 
    ELSIF ((x0 = FALSE) AND  (t0.Q = TRUE) AND  (t1.Q = TRUE)) THEN 
        cstate16 := 27732; y0 := FALSE; y1 := FALSE; y2 := FALSE; t0_start := FALSE;t1_start := TRUE; t1_up := FALSE; 
    ELSIF ((x0 = TRUE) AND  (t0.Q = FALSE) AND  (t1.Q = FALSE)) THEN 
        cstate16 := 48650; y0 := TRUE; y1 := TRUE; y2 := TRUE; t0_start := FALSE;t1_start := FALSE; 
    ELSIF ((x0 = TRUE) AND  (t0.Q = FALSE) AND  (t1.Q = TRUE)) THEN 
        cstate16 := 48646; y0 := TRUE; y1 := TRUE; y2 := TRUE; t0_start := FALSE;t1_start := FALSE; 
    ELSIF ((x0 = TRUE) AND  (t0.Q = TRUE) AND  (t1.Q = FALSE)) THEN 
        cstate16 := 42457; y0 := TRUE; y1 := TRUE; y2 := TRUE; t0_start := FALSE;t1_start := TRUE; t1_up := FALSE; 
    ELSIF ((x0 = TRUE) AND  (t0.Q = TRUE) AND  (t1.Q = TRUE)) THEN 
        cstate16 := 42453; y0 := TRUE; y1 := TRUE; y2 := TRUE; t0_start := FALSE;t1_start := TRUE; t1_up := FALSE; 
    END_IF;
43530:
    IF ((x0 = FALSE) AND  (t0.Q = FALSE) AND  (t1.Q = FALSE)) THEN 
        cstate16 := 34931; y0 := FALSE; y1 := FALSE; y2 := FALSE; t0_start := FALSE;t1_start := FALSE; 
    ELSIF ((x0 = FALSE) AND  (t0.Q = FALSE) AND  (t1.Q = TRUE)) THEN 
        cstate16 := 34932; y0 := FALSE; y1 := FALSE; y2 := FALSE; t0_start := FALSE;t1_start := FALSE; 
    ELSIF ((x0 = FALSE) AND  (t0.Q = TRUE) AND  (t1.Q = FALSE)) THEN 
        cstate16 := 28787; y0 := FALSE; y1 := FALSE; y2 := FALSE; t0_start := FALSE;t1_start := FALSE; 
    ELSIF ((x0 = FALSE) AND  (t0.Q = TRUE) AND  (t1.Q = TRUE)) THEN 
        cstate16 := 28788; y0 := FALSE; y1 := FALSE; y2 := FALSE; t0_start := FALSE;t1_start := FALSE; 
    ELSIF ((x0 = TRUE) AND  (t0.Q = FALSE) AND  (t1.Q = FALSE)) THEN 
        cstate16 := 48650; y0 := TRUE; y1 := TRUE; y2 := TRUE; t0_start := FALSE;t1_start := FALSE; 
    ELSIF ((x0 = TRUE) AND  (t0.Q = FALSE) AND  (t1.Q = TRUE)) THEN 
        cstate16 := 48646; y0 := TRUE; y1 := TRUE; y2 := TRUE; t0_start := FALSE;t1_start := FALSE; 
    ELSIF ((x0 = TRUE) AND  (t0.Q = TRUE) AND  (t1.Q = FALSE)) THEN 
        cstate16 := 43530; y0 := TRUE; y1 := TRUE; y2 := TRUE; t0_start := FALSE;t1_start := FALSE; 
    ELSIF ((x0 = TRUE) AND  (t0.Q = TRUE) AND  (t1.Q = TRUE)) THEN 
        cstate16 := 43526; y0 := TRUE; y1 := TRUE; y2 := TRUE; t0_start := FALSE;t1_start := FALSE; 
    END_IF;
14682:
    IF ((x0 = FALSE) AND  (t0.Q = FALSE) AND  (t1.Q = FALSE)) THEN 
        cstate16 := 34931; y0 := FALSE; y1 := FALSE; y2 := FALSE; t0_start := FALSE;t1_start := FALSE; 
    ELSIF ((x0 = FALSE) AND  (t0.Q = FALSE) AND  (t1.Q = TRUE)) THEN 
        cstate16 := 34932; y0 := FALSE; y1 := FALSE; y2 := FALSE; t0_start := FALSE;t1_start := FALSE; 
    ELSIF ((x0 = FALSE) AND  (t0.Q = TRUE) AND  (t1.Q = FALSE)) THEN 
        cstate16 := 27731; y0 := FALSE; y1 := FALSE; y2 := FALSE; t0_start := FALSE;t1_start := TRUE; t1_up := FALSE; 
    ELSIF ((x0 = FALSE) AND  (t0.Q = TRUE) AND  (t1.Q = TRUE)) THEN 
        cstate16 := 27732; y0 := FALSE; y1 := FALSE; y2 := FALSE; t0_start := FALSE;t1_start := TRUE; t1_up := FALSE; 
    ELSIF ((x0 = TRUE) AND  (t0.Q = FALSE) AND  (t1.Q = FALSE)) THEN 
        cstate16 := 14682; y0 := FALSE; y1 := TRUE; y2 := TRUE; t0_start := FALSE;t1_start := FALSE; 
    ELSIF ((x0 = TRUE) AND  (t0.Q = FALSE) AND  (t1.Q = TRUE)) THEN 
        cstate16 := 14678; y0 := FALSE; y1 := TRUE; y2 := TRUE; t0_start := FALSE;t1_start := FALSE; 
    ELSIF ((x0 = TRUE) AND  (t0.Q = TRUE) AND  (t1.Q = FALSE)) THEN 
        cstate16 := 8361; y0 := FALSE; y1 := TRUE; y2 := TRUE; t0_start := FALSE;t1_start := TRUE; t1_up := FALSE; 
    ELSIF ((x0 = TRUE) AND  (t0.Q = TRUE) AND  (t1.Q = TRUE)) THEN 
        cstate16 := 8357; y0 := FALSE; y1 := TRUE; y2 := TRUE; t0_start := FALSE;t1_start := TRUE; t1_up := FALSE; 
    END_IF;
16689:
    IF ((x0 = FALSE) AND  (t0.Q = FALSE) AND  (t1.Q = FALSE)) THEN 
        cstate16 := 32883; y0 := FALSE; y1 := FALSE; y2 := FALSE; t0_start := FALSE;t1_start := FALSE; 
    ELSIF ((x0 = FALSE) AND  (t0.Q = FALSE) AND  (t1.Q = TRUE)) THEN 
        cstate16 := 34932; y0 := FALSE; y1 := FALSE; y2 := FALSE; t0_start := FALSE;t1_start := FALSE; 
    ELSIF ((x0 = FALSE) AND  (t0.Q = TRUE) AND  (t1.Q = FALSE)) THEN 
        cstate16 := 27731; y0 := FALSE; y1 := FALSE; y2 := FALSE; t0_start := FALSE;t1_start := TRUE; t1_up := FALSE; 
    ELSIF ((x0 = FALSE) AND  (t0.Q = TRUE) AND  (t1.Q = TRUE)) THEN 
        cstate16 := 27732; y0 := FALSE; y1 := FALSE; y2 := FALSE; t0_start := FALSE;t1_start := TRUE; t1_up := FALSE; 
    ELSIF ((x0 = TRUE) AND  (t0.Q = FALSE) AND  (t1.Q = FALSE)) THEN 
        cstate16 := 16689; y0 := FALSE; y1 := TRUE; y2 := FALSE; t0_start := FALSE;t1_start := FALSE; 
    ELSIF ((x0 = TRUE) AND  (t0.Q = FALSE) AND  (t1.Q = TRUE)) THEN 
        cstate16 := 14678; y0 := FALSE; y1 := TRUE; y2 := TRUE; t0_start := FALSE;t1_start := FALSE; 
    ELSIF ((x0 = TRUE) AND  (t0.Q = TRUE) AND  (t1.Q = FALSE)) THEN 
        cstate16 := 8353; y0 := FALSE; y1 := TRUE; y2 := FALSE; t0_start := FALSE;t1_start := TRUE; t1_up := FALSE; 
    ELSIF ((x0 = TRUE) AND  (t0.Q = TRUE) AND  (t1.Q = TRUE)) THEN 
        cstate16 := 8357; y0 := FALSE; y1 := TRUE; y2 := TRUE; t0_start := FALSE;t1_start := TRUE; t1_up := FALSE; 
    END_IF;
48642:
    IF ((x0 = FALSE) AND  (t0.Q = FALSE) AND  (t1.Q = FALSE)) THEN 
        cstate16 := 34931; y0 := FALSE; y1 := FALSE; y2 := FALSE; t0_start := FALSE;t1_start := FALSE; 
    ELSIF ((x0 = FALSE) AND  (t0.Q = FALSE) AND  (t1.Q = TRUE)) THEN 
        cstate16 := 34932; y0 := FALSE; y1 := FALSE; y2 := FALSE; t0_start := FALSE;t1_start := FALSE; 
    ELSIF ((x0 = FALSE) AND  (t0.Q = TRUE) AND  (t1.Q = FALSE)) THEN 
        cstate16 := 27731; y0 := FALSE; y1 := FALSE; y2 := FALSE; t0_start := FALSE;t1_start := TRUE; t1_up := FALSE; 
    ELSIF ((x0 = FALSE) AND  (t0.Q = TRUE) AND  (t1.Q = TRUE)) THEN 
        cstate16 := 27732; y0 := FALSE; y1 := FALSE; y2 := FALSE; t0_start := FALSE;t1_start := TRUE; t1_up := FALSE; 
    ELSIF ((x0 = TRUE) AND  (t0.Q = FALSE) AND  (t1.Q = FALSE)) THEN 
        cstate16 := 48641; y0 := TRUE; y1 := TRUE; y2 := FALSE; t0_start := FALSE;t1_start := FALSE; 
    ELSIF ((x0 = TRUE) AND  (t0.Q = FALSE) AND  (t1.Q = TRUE)) THEN 
        cstate16 := 48642; y0 := TRUE; y1 := TRUE; y2 := FALSE; t0_start := FALSE;t1_start := FALSE; 
    ELSIF ((x0 = TRUE) AND  (t0.Q = TRUE) AND  (t1.Q = FALSE)) THEN 
        cstate16 := 42449; y0 := TRUE; y1 := TRUE; y2 := FALSE; t0_start := FALSE;t1_start := TRUE; t1_up := FALSE; 
    ELSIF ((x0 = TRUE) AND  (t0.Q = TRUE) AND  (t1.Q = TRUE)) THEN 
        cstate16 := 42450; y0 := TRUE; y1 := TRUE; y2 := FALSE; t0_start := FALSE;t1_start := TRUE; t1_up := FALSE; 
    END_IF;
14674:
    IF ((x0 = FALSE) AND  (t0.Q = FALSE) AND  (t1.Q = FALSE)) THEN 
        cstate16 := 34931; y0 := FALSE; y1 := FALSE; y2 := FALSE; t0_start := FALSE;t1_start := FALSE; 
    ELSIF ((x0 = FALSE) AND  (t0.Q = FALSE) AND  (t1.Q = TRUE)) THEN 
        cstate16 := 34932; y0 := FALSE; y1 := FALSE; y2 := FALSE; t0_start := FALSE;t1_start := FALSE; 
    ELSIF ((x0 = FALSE) AND  (t0.Q = TRUE) AND  (t1.Q = FALSE)) THEN 
        cstate16 := 27731; y0 := FALSE; y1 := FALSE; y2 := FALSE; t0_start := FALSE;t1_start := TRUE; t1_up := FALSE; 
    ELSIF ((x0 = FALSE) AND  (t0.Q = TRUE) AND  (t1.Q = TRUE)) THEN 
        cstate16 := 27732; y0 := FALSE; y1 := FALSE; y2 := FALSE; t0_start := FALSE;t1_start := TRUE; t1_up := FALSE; 
    ELSIF ((x0 = TRUE) AND  (t0.Q = FALSE) AND  (t1.Q = FALSE)) THEN 
        cstate16 := 14673; y0 := FALSE; y1 := TRUE; y2 := FALSE; t0_start := FALSE;t1_start := FALSE; 
    ELSIF ((x0 = TRUE) AND  (t0.Q = FALSE) AND  (t1.Q = TRUE)) THEN 
        cstate16 := 14674; y0 := FALSE; y1 := TRUE; y2 := FALSE; t0_start := FALSE;t1_start := FALSE; 
    ELSIF ((x0 = TRUE) AND  (t0.Q = TRUE) AND  (t1.Q = FALSE)) THEN 
        cstate16 := 8353; y0 := FALSE; y1 := TRUE; y2 := FALSE; t0_start := FALSE;t1_start := TRUE; t1_up := FALSE; 
    ELSIF ((x0 = TRUE) AND  (t0.Q = TRUE) AND  (t1.Q = TRUE)) THEN 
        cstate16 := 8354; y0 := FALSE; y1 := TRUE; y2 := FALSE; t0_start := FALSE;t1_start := TRUE; t1_up := FALSE; 
    END_IF;
47799:
    IF ((x0 = FALSE) AND  (t0.Q = FALSE) AND  (t1.Q = FALSE)) THEN 
        cstate16 := 34931; y0 := FALSE; y1 := FALSE; y2 := FALSE; t0_start := FALSE;t1_start := FALSE; 
    ELSIF ((x0 = FALSE) AND  (t0.Q = FALSE) AND  (t1.Q = TRUE)) THEN 
        cstate16 := 34932; y0 := FALSE; y1 := FALSE; y2 := FALSE; t0_start := FALSE;t1_start := FALSE; 
    ELSIF ((x0 = FALSE) AND  (t0.Q = TRUE) AND  (t1.Q = FALSE)) THEN 
        cstate16 := 28787; y0 := FALSE; y1 := FALSE; y2 := FALSE; t0_start := FALSE;t1_start := FALSE; 
    ELSIF ((x0 = FALSE) AND  (t0.Q = TRUE) AND  (t1.Q = TRUE)) THEN 
        cstate16 := 28788; y0 := FALSE; y1 := FALSE; y2 := FALSE; t0_start := FALSE;t1_start := FALSE; 
    ELSIF ((x0 = TRUE) AND  (t0.Q = FALSE) AND  (t1.Q = FALSE)) THEN 
        cstate16 := 40652; y0 := TRUE; y1 := TRUE; y2 := TRUE; t0_start := TRUE; t0_up := FALSE;t1_start := FALSE; 
    ELSIF ((x0 = TRUE) AND  (t0.Q = FALSE) AND  (t1.Q = TRUE)) THEN 
        cstate16 := 40647; y0 := TRUE; y1 := TRUE; y2 := TRUE; t0_start := TRUE; t0_up := FALSE;t1_start := FALSE; 
    ELSIF ((x0 = TRUE) AND  (t0.Q = TRUE) AND  (t1.Q = FALSE)) THEN 
        cstate16 := 47804; y0 := TRUE; y1 := TRUE; y2 := TRUE; t0_start := FALSE;t1_start := FALSE; 
    ELSIF ((x0 = TRUE) AND  (t0.Q = TRUE) AND  (t1.Q = TRUE)) THEN 
        cstate16 := 47799; y0 := TRUE; y1 := TRUE; y2 := TRUE; t0_start := FALSE;t1_start := FALSE; 
    END_IF;
43410:
    IF ((x0 = FALSE) AND  (t0.Q = FALSE) AND  (t1.Q = FALSE)) THEN 
        cstate16 := 34931; y0 := FALSE; y1 := FALSE; y2 := FALSE; t0_start := FALSE;t1_start := FALSE; 
    ELSIF ((x0 = FALSE) AND  (t0.Q = FALSE) AND  (t1.Q = TRUE)) THEN 
        cstate16 := 34932; y0 := FALSE; y1 := FALSE; y2 := FALSE; t0_start := FALSE;t1_start := FALSE; 
    ELSIF ((x0 = FALSE) AND  (t0.Q = TRUE) AND  (t1.Q = FALSE)) THEN 
        cstate16 := 28787; y0 := FALSE; y1 := FALSE; y2 := FALSE; t0_start := FALSE;t1_start := FALSE; 
    ELSIF ((x0 = FALSE) AND  (t0.Q = TRUE) AND  (t1.Q = TRUE)) THEN 
        cstate16 := 28788; y0 := FALSE; y1 := FALSE; y2 := FALSE; t0_start := FALSE;t1_start := FALSE; 
    ELSIF ((x0 = TRUE) AND  (t0.Q = FALSE) AND  (t1.Q = FALSE)) THEN 
        cstate16 := 48529; y0 := TRUE; y1 := FALSE; y2 := FALSE; t0_start := FALSE;t1_start := FALSE; 
    ELSIF ((x0 = TRUE) AND  (t0.Q = FALSE) AND  (t1.Q = TRUE)) THEN 
        cstate16 := 48530; y0 := TRUE; y1 := FALSE; y2 := FALSE; t0_start := FALSE;t1_start := FALSE; 
    ELSIF ((x0 = TRUE) AND  (t0.Q = TRUE) AND  (t1.Q = FALSE)) THEN 
        cstate16 := 43409; y0 := TRUE; y1 := FALSE; y2 := FALSE; t0_start := FALSE;t1_start := FALSE; 
    ELSIF ((x0 = TRUE) AND  (t0.Q = TRUE) AND  (t1.Q = TRUE)) THEN 
        cstate16 := 43410; y0 := TRUE; y1 := FALSE; y2 := FALSE; t0_start := FALSE;t1_start := FALSE; 
    END_IF;
25129:
    IF ((x0 = FALSE) AND  (t0.Q = FALSE) AND  (t1.Q = FALSE)) THEN 
        cstate16 := 23667; y0 := FALSE; y1 := FALSE; y2 := FALSE; t0_start := FALSE;t1_start := FALSE; 
    ELSIF ((x0 = FALSE) AND  (t0.Q = FALSE) AND  (t1.Q = TRUE)) THEN 
        cstate16 := 26740; y0 := FALSE; y1 := FALSE; y2 := FALSE; t0_start := FALSE;t1_start := FALSE; 
    ELSIF ((x0 = FALSE) AND  (t0.Q = TRUE) AND  (t1.Q = FALSE)) THEN 
        cstate16 := 17491; y0 := FALSE; y1 := FALSE; y2 := FALSE; t0_start := FALSE;t1_start := TRUE; t1_up := FALSE; 
    ELSIF ((x0 = FALSE) AND  (t0.Q = TRUE) AND  (t1.Q = TRUE)) THEN 
        cstate16 := 17492; y0 := FALSE; y1 := FALSE; y2 := FALSE; t0_start := FALSE;t1_start := TRUE; t1_up := FALSE; 
    ELSIF ((x0 = TRUE) AND  (t0.Q = FALSE) AND  (t1.Q = FALSE)) THEN 
        cstate16 := 25129; y0 := TRUE; y1 := TRUE; y2 := TRUE; t0_start := FALSE;t1_start := FALSE; 
    ELSIF ((x0 = TRUE) AND  (t0.Q = FALSE) AND  (t1.Q = TRUE)) THEN 
        cstate16 := 26134; y0 := TRUE; y1 := TRUE; y2 := TRUE; t0_start := FALSE;t1_start := FALSE; 
    ELSIF ((x0 = TRUE) AND  (t0.Q = TRUE) AND  (t1.Q = FALSE)) THEN 
        cstate16 := 42457; y0 := TRUE; y1 := TRUE; y2 := TRUE; t0_start := FALSE;t1_start := TRUE; t1_up := FALSE; 
    ELSIF ((x0 = TRUE) AND  (t0.Q = TRUE) AND  (t1.Q = TRUE)) THEN 
        cstate16 := 42453; y0 := TRUE; y1 := TRUE; y2 := TRUE; t0_start := FALSE;t1_start := TRUE; t1_up := FALSE; 
    END_IF;
38147:
    IF ((x0 = FALSE) AND  (t0.Q = FALSE) AND  (t1.Q = FALSE)) THEN 
        cstate16 := 23667; y0 := FALSE; y1 := FALSE; y2 := FALSE; t0_start := FALSE;t1_start := FALSE; 
    ELSIF ((x0 = FALSE) AND  (t0.Q = FALSE) AND  (t1.Q = TRUE)) THEN 
        cstate16 := 26740; y0 := FALSE; y1 := FALSE; y2 := FALSE; t0_start := FALSE;t1_start := FALSE; 
    ELSIF ((x0 = FALSE) AND  (t0.Q = TRUE) AND  (t1.Q = FALSE)) THEN 
        cstate16 := 17523; y0 := FALSE; y1 := FALSE; y2 := FALSE; t0_start := FALSE;t1_start := FALSE; 
    ELSIF ((x0 = FALSE) AND  (t0.Q = TRUE) AND  (t1.Q = TRUE)) THEN 
        cstate16 := 22644; y0 := FALSE; y1 := FALSE; y2 := FALSE; t0_start := FALSE;t1_start := FALSE; 
    ELSIF ((x0 = TRUE) AND  (t0.Q = FALSE) AND  (t1.Q = FALSE)) THEN 
        cstate16 := 41699; y0 := TRUE; y1 := TRUE; y2 := FALSE; t0_start := FALSE;t1_start := FALSE; 
    ELSIF ((x0 = TRUE) AND  (t0.Q = FALSE) AND  (t1.Q = TRUE)) THEN 
        cstate16 := 40663; y0 := TRUE; y1 := TRUE; y2 := TRUE; t0_start := FALSE;t1_start := FALSE; 
    ELSIF ((x0 = TRUE) AND  (t0.Q = TRUE) AND  (t1.Q = FALSE)) THEN 
        cstate16 := 46739; y0 := TRUE; y1 := TRUE; y2 := FALSE; t0_start := FALSE;t1_start := FALSE; 
    ELSIF ((x0 = TRUE) AND  (t0.Q = TRUE) AND  (t1.Q = TRUE)) THEN 
        cstate16 := 47799; y0 := TRUE; y1 := TRUE; y2 := TRUE; t0_start := FALSE;t1_start := FALSE; 
    END_IF;
32883:
    IF ((x0 = FALSE) AND  (t0.Q = FALSE) AND  (t1.Q = FALSE)) THEN 
        cstate16 := 32883; y0 := FALSE; y1 := FALSE; y2 := FALSE; t0_start := FALSE;t1_start := FALSE; 
    ELSIF ((x0 = FALSE) AND  (t0.Q = FALSE) AND  (t1.Q = TRUE)) THEN 
        cstate16 := 34932; y0 := FALSE; y1 := FALSE; y2 := FALSE; t0_start := FALSE;t1_start := FALSE; 
    ELSIF ((x0 = FALSE) AND  (t0.Q = TRUE) AND  (t1.Q = FALSE)) THEN 
        cstate16 := 27731; y0 := FALSE; y1 := FALSE; y2 := FALSE; t0_start := FALSE;t1_start := TRUE; t1_up := FALSE; 
    ELSIF ((x0 = FALSE) AND  (t0.Q = TRUE) AND  (t1.Q = TRUE)) THEN 
        cstate16 := 27732; y0 := FALSE; y1 := FALSE; y2 := FALSE; t0_start := FALSE;t1_start := TRUE; t1_up := FALSE; 
    ELSIF ((x0 = TRUE) AND  (t0.Q = FALSE) AND  (t1.Q = FALSE)) THEN 
        cstate16 := 41187; y0 := TRUE; y1 := FALSE; y2 := FALSE; t0_start := TRUE; t0_up := FALSE;t1_start := FALSE; 
    ELSIF ((x0 = TRUE) AND  (t0.Q = FALSE) AND  (t1.Q = TRUE)) THEN 
        cstate16 := 40167; y0 := TRUE; y1 := FALSE; y2 := TRUE; t0_start := TRUE; t0_up := FALSE;t1_start := FALSE; 
    ELSIF ((x0 = TRUE) AND  (t0.Q = TRUE) AND  (t1.Q = FALSE)) THEN 
        cstate16 := 38147; y0 := TRUE; y1 := TRUE; y2 := FALSE; t0_start := TRUE; t0_up := FALSE;t1_start := TRUE; t1_up := FALSE; 
    ELSIF ((x0 = TRUE) AND  (t0.Q = TRUE) AND  (t1.Q = TRUE)) THEN 
        cstate16 := 38152; y0 := TRUE; y1 := TRUE; y2 := TRUE; t0_start := TRUE; t0_up := FALSE;t1_start := TRUE; t1_up := FALSE; 
    END_IF;
47796:
    IF ((x0 = FALSE) AND  (t0.Q = FALSE) AND  (t1.Q = FALSE)) THEN 
        cstate16 := 34931; y0 := FALSE; y1 := FALSE; y2 := FALSE; t0_start := FALSE;t1_start := FALSE; 
    ELSIF ((x0 = FALSE) AND  (t0.Q = FALSE) AND  (t1.Q = TRUE)) THEN 
        cstate16 := 34932; y0 := FALSE; y1 := FALSE; y2 := FALSE; t0_start := FALSE;t1_start := FALSE; 
    ELSIF ((x0 = FALSE) AND  (t0.Q = TRUE) AND  (t1.Q = FALSE)) THEN 
        cstate16 := 28787; y0 := FALSE; y1 := FALSE; y2 := FALSE; t0_start := FALSE;t1_start := FALSE; 
    ELSIF ((x0 = FALSE) AND  (t0.Q = TRUE) AND  (t1.Q = TRUE)) THEN 
        cstate16 := 28788; y0 := FALSE; y1 := FALSE; y2 := FALSE; t0_start := FALSE;t1_start := FALSE; 
    ELSIF ((x0 = TRUE) AND  (t0.Q = FALSE) AND  (t1.Q = FALSE)) THEN 
        cstate16 := 40643; y0 := TRUE; y1 := TRUE; y2 := FALSE; t0_start := TRUE; t0_up := FALSE;t1_start := FALSE; 
    ELSIF ((x0 = TRUE) AND  (t0.Q = FALSE) AND  (t1.Q = TRUE)) THEN 
        cstate16 := 40644; y0 := TRUE; y1 := TRUE; y2 := FALSE; t0_start := TRUE; t0_up := FALSE;t1_start := FALSE; 
    ELSIF ((x0 = TRUE) AND  (t0.Q = TRUE) AND  (t1.Q = FALSE)) THEN 
        cstate16 := 47795; y0 := TRUE; y1 := TRUE; y2 := FALSE; t0_start := FALSE;t1_start := FALSE; 
    ELSIF ((x0 = TRUE) AND  (t0.Q = TRUE) AND  (t1.Q = TRUE)) THEN 
        cstate16 := 47796; y0 := TRUE; y1 := TRUE; y2 := FALSE; t0_start := FALSE;t1_start := FALSE; 
    END_IF;
14678:
    IF ((x0 = FALSE) AND  (t0.Q = FALSE) AND  (t1.Q = FALSE)) THEN 
        cstate16 := 34931; y0 := FALSE; y1 := FALSE; y2 := FALSE; t0_start := FALSE;t1_start := FALSE; 
    ELSIF ((x0 = FALSE) AND  (t0.Q = FALSE) AND  (t1.Q = TRUE)) THEN 
        cstate16 := 34932; y0 := FALSE; y1 := FALSE; y2 := FALSE; t0_start := FALSE;t1_start := FALSE; 
    ELSIF ((x0 = FALSE) AND  (t0.Q = TRUE) AND  (t1.Q = FALSE)) THEN 
        cstate16 := 27731; y0 := FALSE; y1 := FALSE; y2 := FALSE; t0_start := FALSE;t1_start := TRUE; t1_up := FALSE; 
    ELSIF ((x0 = FALSE) AND  (t0.Q = TRUE) AND  (t1.Q = TRUE)) THEN 
        cstate16 := 27732; y0 := FALSE; y1 := FALSE; y2 := FALSE; t0_start := FALSE;t1_start := TRUE; t1_up := FALSE; 
    ELSIF ((x0 = TRUE) AND  (t0.Q = FALSE) AND  (t1.Q = FALSE)) THEN 
        cstate16 := 14682; y0 := FALSE; y1 := TRUE; y2 := TRUE; t0_start := FALSE;t1_start := FALSE; 
    ELSIF ((x0 = TRUE) AND  (t0.Q = FALSE) AND  (t1.Q = TRUE)) THEN 
        cstate16 := 14678; y0 := FALSE; y1 := TRUE; y2 := TRUE; t0_start := FALSE;t1_start := FALSE; 
    ELSIF ((x0 = TRUE) AND  (t0.Q = TRUE) AND  (t1.Q = FALSE)) THEN 
        cstate16 := 8361; y0 := FALSE; y1 := TRUE; y2 := TRUE; t0_start := FALSE;t1_start := TRUE; t1_up := FALSE; 
    ELSIF ((x0 = TRUE) AND  (t0.Q = TRUE) AND  (t1.Q = TRUE)) THEN 
        cstate16 := 8357; y0 := FALSE; y1 := TRUE; y2 := TRUE; t0_start := FALSE;t1_start := TRUE; t1_up := FALSE; 
    END_IF;
47795:
    IF ((x0 = FALSE) AND  (t0.Q = FALSE) AND  (t1.Q = FALSE)) THEN 
        cstate16 := 34931; y0 := FALSE; y1 := FALSE; y2 := FALSE; t0_start := FALSE;t1_start := FALSE; 
    ELSIF ((x0 = FALSE) AND  (t0.Q = FALSE) AND  (t1.Q = TRUE)) THEN 
        cstate16 := 34932; y0 := FALSE; y1 := FALSE; y2 := FALSE; t0_start := FALSE;t1_start := FALSE; 
    ELSIF ((x0 = FALSE) AND  (t0.Q = TRUE) AND  (t1.Q = FALSE)) THEN 
        cstate16 := 28787; y0 := FALSE; y1 := FALSE; y2 := FALSE; t0_start := FALSE;t1_start := FALSE; 
    ELSIF ((x0 = FALSE) AND  (t0.Q = TRUE) AND  (t1.Q = TRUE)) THEN 
        cstate16 := 28788; y0 := FALSE; y1 := FALSE; y2 := FALSE; t0_start := FALSE;t1_start := FALSE; 
    ELSIF ((x0 = TRUE) AND  (t0.Q = FALSE) AND  (t1.Q = FALSE)) THEN 
        cstate16 := 40643; y0 := TRUE; y1 := TRUE; y2 := FALSE; t0_start := TRUE; t0_up := FALSE;t1_start := FALSE; 
    ELSIF ((x0 = TRUE) AND  (t0.Q = FALSE) AND  (t1.Q = TRUE)) THEN 
        cstate16 := 40647; y0 := TRUE; y1 := TRUE; y2 := TRUE; t0_start := TRUE; t0_up := FALSE;t1_start := FALSE; 
    ELSIF ((x0 = TRUE) AND  (t0.Q = TRUE) AND  (t1.Q = FALSE)) THEN 
        cstate16 := 47795; y0 := TRUE; y1 := TRUE; y2 := FALSE; t0_start := FALSE;t1_start := FALSE; 
    ELSIF ((x0 = TRUE) AND  (t0.Q = TRUE) AND  (t1.Q = TRUE)) THEN 
        cstate16 := 47799; y0 := TRUE; y1 := TRUE; y2 := TRUE; t0_start := FALSE;t1_start := FALSE; 
    END_IF;
6218:
    IF ((x0 = FALSE) AND  (t0.Q = FALSE) AND  (t1.Q = FALSE)) THEN 
        cstate16 := 34931; y0 := FALSE; y1 := FALSE; y2 := FALSE; t0_start := FALSE;t1_start := FALSE; 
    ELSIF ((x0 = FALSE) AND  (t0.Q = FALSE) AND  (t1.Q = TRUE)) THEN 
        cstate16 := 34932; y0 := FALSE; y1 := FALSE; y2 := FALSE; t0_start := FALSE;t1_start := FALSE; 
    ELSIF ((x0 = FALSE) AND  (t0.Q = TRUE) AND  (t1.Q = FALSE)) THEN 
        cstate16 := 28787; y0 := FALSE; y1 := FALSE; y2 := FALSE; t0_start := FALSE;t1_start := FALSE; 
    ELSIF ((x0 = FALSE) AND  (t0.Q = TRUE) AND  (t1.Q = TRUE)) THEN 
        cstate16 := 28788; y0 := FALSE; y1 := FALSE; y2 := FALSE; t0_start := FALSE;t1_start := FALSE; 
    ELSIF ((x0 = TRUE) AND  (t0.Q = FALSE) AND  (t1.Q = FALSE)) THEN 
        cstate16 := 14410; y0 := FALSE; y1 := FALSE; y2 := TRUE; t0_start := FALSE;t1_start := FALSE; 
    ELSIF ((x0 = TRUE) AND  (t0.Q = FALSE) AND  (t1.Q = TRUE)) THEN 
        cstate16 := 14406; y0 := FALSE; y1 := FALSE; y2 := TRUE; t0_start := FALSE;t1_start := FALSE; 
    ELSIF ((x0 = TRUE) AND  (t0.Q = TRUE) AND  (t1.Q = FALSE)) THEN 
        cstate16 := 6218; y0 := FALSE; y1 := FALSE; y2 := TRUE; t0_start := FALSE;t1_start := FALSE; 
    ELSIF ((x0 = TRUE) AND  (t0.Q = TRUE) AND  (t1.Q = TRUE)) THEN 
        cstate16 := 6214; y0 := FALSE; y1 := FALSE; y2 := TRUE; t0_start := FALSE;t1_start := FALSE; 
    END_IF;
17492:
    IF ((x0 = FALSE) AND  (t0.Q = FALSE) AND  (t1.Q = FALSE)) THEN 
        cstate16 := 32883; y0 := FALSE; y1 := FALSE; y2 := FALSE; t0_start := FALSE;t1_start := FALSE; 
    ELSIF ((x0 = FALSE) AND  (t0.Q = FALSE) AND  (t1.Q = TRUE)) THEN 
        cstate16 := 34932; y0 := FALSE; y1 := FALSE; y2 := FALSE; t0_start := FALSE;t1_start := FALSE; 
    ELSIF ((x0 = FALSE) AND  (t0.Q = TRUE) AND  (t1.Q = FALSE)) THEN 
        cstate16 := 27763; y0 := FALSE; y1 := FALSE; y2 := FALSE; t0_start := FALSE;t1_start := FALSE; 
    ELSIF ((x0 = FALSE) AND  (t0.Q = TRUE) AND  (t1.Q = TRUE)) THEN 
        cstate16 := 28788; y0 := FALSE; y1 := FALSE; y2 := FALSE; t0_start := FALSE;t1_start := FALSE; 
    ELSIF ((x0 = TRUE) AND  (t0.Q = FALSE) AND  (t1.Q = FALSE)) THEN 
        cstate16 := 41187; y0 := TRUE; y1 := FALSE; y2 := FALSE; t0_start := TRUE; t0_up := FALSE;t1_start := FALSE; 
    ELSIF ((x0 = TRUE) AND  (t0.Q = FALSE) AND  (t1.Q = TRUE)) THEN 
        cstate16 := 40164; y0 := TRUE; y1 := FALSE; y2 := FALSE; t0_start := TRUE; t0_up := FALSE;t1_start := FALSE; 
    ELSIF ((x0 = TRUE) AND  (t0.Q = TRUE) AND  (t1.Q = FALSE)) THEN 
        cstate16 := 38115; y0 := TRUE; y1 := FALSE; y2 := FALSE; t0_start := TRUE; t0_up := FALSE;t1_start := FALSE; 
    ELSIF ((x0 = TRUE) AND  (t0.Q = TRUE) AND  (t1.Q = TRUE)) THEN 
        cstate16 := 39140; y0 := TRUE; y1 := FALSE; y2 := FALSE; t0_start := TRUE; t0_up := FALSE;t1_start := FALSE; 
    END_IF;
43418:
    IF ((x0 = FALSE) AND  (t0.Q = FALSE) AND  (t1.Q = FALSE)) THEN 
        cstate16 := 34931; y0 := FALSE; y1 := FALSE; y2 := FALSE; t0_start := FALSE;t1_start := FALSE; 
    ELSIF ((x0 = FALSE) AND  (t0.Q = FALSE) AND  (t1.Q = TRUE)) THEN 
        cstate16 := 34932; y0 := FALSE; y1 := FALSE; y2 := FALSE; t0_start := FALSE;t1_start := FALSE; 
    ELSIF ((x0 = FALSE) AND  (t0.Q = TRUE) AND  (t1.Q = FALSE)) THEN 
        cstate16 := 28787; y0 := FALSE; y1 := FALSE; y2 := FALSE; t0_start := FALSE;t1_start := FALSE; 
    ELSIF ((x0 = FALSE) AND  (t0.Q = TRUE) AND  (t1.Q = TRUE)) THEN 
        cstate16 := 28788; y0 := FALSE; y1 := FALSE; y2 := FALSE; t0_start := FALSE;t1_start := FALSE; 
    ELSIF ((x0 = TRUE) AND  (t0.Q = FALSE) AND  (t1.Q = FALSE)) THEN 
        cstate16 := 48538; y0 := TRUE; y1 := FALSE; y2 := TRUE; t0_start := FALSE;t1_start := FALSE; 
    ELSIF ((x0 = TRUE) AND  (t0.Q = FALSE) AND  (t1.Q = TRUE)) THEN 
        cstate16 := 48534; y0 := TRUE; y1 := FALSE; y2 := TRUE; t0_start := FALSE;t1_start := FALSE; 
    ELSIF ((x0 = TRUE) AND  (t0.Q = TRUE) AND  (t1.Q = FALSE)) THEN 
        cstate16 := 43418; y0 := TRUE; y1 := FALSE; y2 := TRUE; t0_start := FALSE;t1_start := FALSE; 
    ELSIF ((x0 = TRUE) AND  (t0.Q = TRUE) AND  (t1.Q = TRUE)) THEN 
        cstate16 := 43414; y0 := TRUE; y1 := FALSE; y2 := TRUE; t0_start := FALSE;t1_start := FALSE; 
    END_IF;
17491:
    IF ((x0 = FALSE) AND  (t0.Q = FALSE) AND  (t1.Q = FALSE)) THEN 
        cstate16 := 32883; y0 := FALSE; y1 := FALSE; y2 := FALSE; t0_start := FALSE;t1_start := FALSE; 
    ELSIF ((x0 = FALSE) AND  (t0.Q = FALSE) AND  (t1.Q = TRUE)) THEN 
        cstate16 := 34932; y0 := FALSE; y1 := FALSE; y2 := FALSE; t0_start := FALSE;t1_start := FALSE; 
    ELSIF ((x0 = FALSE) AND  (t0.Q = TRUE) AND  (t1.Q = FALSE)) THEN 
        cstate16 := 27763; y0 := FALSE; y1 := FALSE; y2 := FALSE; t0_start := FALSE;t1_start := FALSE; 
    ELSIF ((x0 = FALSE) AND  (t0.Q = TRUE) AND  (t1.Q = TRUE)) THEN 
        cstate16 := 28788; y0 := FALSE; y1 := FALSE; y2 := FALSE; t0_start := FALSE;t1_start := FALSE; 
    ELSIF ((x0 = TRUE) AND  (t0.Q = FALSE) AND  (t1.Q = FALSE)) THEN 
        cstate16 := 41187; y0 := TRUE; y1 := FALSE; y2 := FALSE; t0_start := TRUE; t0_up := FALSE;t1_start := FALSE; 
    ELSIF ((x0 = TRUE) AND  (t0.Q = FALSE) AND  (t1.Q = TRUE)) THEN 
        cstate16 := 40167; y0 := TRUE; y1 := FALSE; y2 := TRUE; t0_start := TRUE; t0_up := FALSE;t1_start := FALSE; 
    ELSIF ((x0 = TRUE) AND  (t0.Q = TRUE) AND  (t1.Q = FALSE)) THEN 
        cstate16 := 38115; y0 := TRUE; y1 := FALSE; y2 := FALSE; t0_start := TRUE; t0_up := FALSE;t1_start := FALSE; 
    ELSIF ((x0 = TRUE) AND  (t0.Q = TRUE) AND  (t1.Q = TRUE)) THEN 
        cstate16 := 39143; y0 := TRUE; y1 := FALSE; y2 := TRUE; t0_start := TRUE; t0_up := FALSE;t1_start := FALSE; 
    END_IF;
48530:
    IF ((x0 = FALSE) AND  (t0.Q = FALSE) AND  (t1.Q = FALSE)) THEN 
        cstate16 := 34931; y0 := FALSE; y1 := FALSE; y2 := FALSE; t0_start := FALSE;t1_start := FALSE; 
    ELSIF ((x0 = FALSE) AND  (t0.Q = FALSE) AND  (t1.Q = TRUE)) THEN 
        cstate16 := 34932; y0 := FALSE; y1 := FALSE; y2 := FALSE; t0_start := FALSE;t1_start := FALSE; 
    ELSIF ((x0 = FALSE) AND  (t0.Q = TRUE) AND  (t1.Q = FALSE)) THEN 
        cstate16 := 27731; y0 := FALSE; y1 := FALSE; y2 := FALSE; t0_start := FALSE;t1_start := TRUE; t1_up := FALSE; 
    ELSIF ((x0 = FALSE) AND  (t0.Q = TRUE) AND  (t1.Q = TRUE)) THEN 
        cstate16 := 27732; y0 := FALSE; y1 := FALSE; y2 := FALSE; t0_start := FALSE;t1_start := TRUE; t1_up := FALSE; 
    ELSIF ((x0 = TRUE) AND  (t0.Q = FALSE) AND  (t1.Q = FALSE)) THEN 
        cstate16 := 48529; y0 := TRUE; y1 := FALSE; y2 := FALSE; t0_start := FALSE;t1_start := FALSE; 
    ELSIF ((x0 = TRUE) AND  (t0.Q = FALSE) AND  (t1.Q = TRUE)) THEN 
        cstate16 := 48530; y0 := TRUE; y1 := FALSE; y2 := FALSE; t0_start := FALSE;t1_start := FALSE; 
    ELSIF ((x0 = TRUE) AND  (t0.Q = TRUE) AND  (t1.Q = FALSE)) THEN 
        cstate16 := 42449; y0 := TRUE; y1 := TRUE; y2 := FALSE; t0_start := FALSE;t1_start := TRUE; t1_up := FALSE; 
    ELSIF ((x0 = TRUE) AND  (t0.Q = TRUE) AND  (t1.Q = TRUE)) THEN 
        cstate16 := 42450; y0 := TRUE; y1 := TRUE; y2 := FALSE; t0_start := FALSE;t1_start := TRUE; t1_up := FALSE; 
    END_IF;
8497:
    IF ((x0 = FALSE) AND  (t0.Q = FALSE) AND  (t1.Q = FALSE)) THEN 
        cstate16 := 32883; y0 := FALSE; y1 := FALSE; y2 := FALSE; t0_start := FALSE;t1_start := FALSE; 
    ELSIF ((x0 = FALSE) AND  (t0.Q = FALSE) AND  (t1.Q = TRUE)) THEN 
        cstate16 := 34932; y0 := FALSE; y1 := FALSE; y2 := FALSE; t0_start := FALSE;t1_start := FALSE; 
    ELSIF ((x0 = FALSE) AND  (t0.Q = TRUE) AND  (t1.Q = FALSE)) THEN 
        cstate16 := 27763; y0 := FALSE; y1 := FALSE; y2 := FALSE; t0_start := FALSE;t1_start := FALSE; 
    ELSIF ((x0 = FALSE) AND  (t0.Q = TRUE) AND  (t1.Q = TRUE)) THEN 
        cstate16 := 28788; y0 := FALSE; y1 := FALSE; y2 := FALSE; t0_start := FALSE;t1_start := FALSE; 
    ELSIF ((x0 = TRUE) AND  (t0.Q = FALSE) AND  (t1.Q = FALSE)) THEN 
        cstate16 := 16689; y0 := FALSE; y1 := TRUE; y2 := FALSE; t0_start := FALSE;t1_start := FALSE; 
    ELSIF ((x0 = TRUE) AND  (t0.Q = FALSE) AND  (t1.Q = TRUE)) THEN 
        cstate16 := 14678; y0 := FALSE; y1 := TRUE; y2 := TRUE; t0_start := FALSE;t1_start := FALSE; 
    ELSIF ((x0 = TRUE) AND  (t0.Q = TRUE) AND  (t1.Q = FALSE)) THEN 
        cstate16 := 8497; y0 := FALSE; y1 := TRUE; y2 := FALSE; t0_start := FALSE;t1_start := FALSE; 
    ELSIF ((x0 = TRUE) AND  (t0.Q = TRUE) AND  (t1.Q = TRUE)) THEN 
        cstate16 := 6486; y0 := FALSE; y1 := TRUE; y2 := TRUE; t0_start := FALSE;t1_start := FALSE; 
    END_IF;
43414:
    IF ((x0 = FALSE) AND  (t0.Q = FALSE) AND  (t1.Q = FALSE)) THEN 
        cstate16 := 34931; y0 := FALSE; y1 := FALSE; y2 := FALSE; t0_start := FALSE;t1_start := FALSE; 
    ELSIF ((x0 = FALSE) AND  (t0.Q = FALSE) AND  (t1.Q = TRUE)) THEN 
        cstate16 := 34932; y0 := FALSE; y1 := FALSE; y2 := FALSE; t0_start := FALSE;t1_start := FALSE; 
    ELSIF ((x0 = FALSE) AND  (t0.Q = TRUE) AND  (t1.Q = FALSE)) THEN 
        cstate16 := 28787; y0 := FALSE; y1 := FALSE; y2 := FALSE; t0_start := FALSE;t1_start := FALSE; 
    ELSIF ((x0 = FALSE) AND  (t0.Q = TRUE) AND  (t1.Q = TRUE)) THEN 
        cstate16 := 28788; y0 := FALSE; y1 := FALSE; y2 := FALSE; t0_start := FALSE;t1_start := FALSE; 
    ELSIF ((x0 = TRUE) AND  (t0.Q = FALSE) AND  (t1.Q = FALSE)) THEN 
        cstate16 := 48538; y0 := TRUE; y1 := FALSE; y2 := TRUE; t0_start := FALSE;t1_start := FALSE; 
    ELSIF ((x0 = TRUE) AND  (t0.Q = FALSE) AND  (t1.Q = TRUE)) THEN 
        cstate16 := 48534; y0 := TRUE; y1 := FALSE; y2 := TRUE; t0_start := FALSE;t1_start := FALSE; 
    ELSIF ((x0 = TRUE) AND  (t0.Q = TRUE) AND  (t1.Q = FALSE)) THEN 
        cstate16 := 43418; y0 := TRUE; y1 := FALSE; y2 := TRUE; t0_start := FALSE;t1_start := FALSE; 
    ELSIF ((x0 = TRUE) AND  (t0.Q = TRUE) AND  (t1.Q = TRUE)) THEN 
        cstate16 := 43414; y0 := TRUE; y1 := FALSE; y2 := TRUE; t0_start := FALSE;t1_start := FALSE; 
    END_IF;
43526:
    IF ((x0 = FALSE) AND  (t0.Q = FALSE) AND  (t1.Q = FALSE)) THEN 
        cstate16 := 34931; y0 := FALSE; y1 := FALSE; y2 := FALSE; t0_start := FALSE;t1_start := FALSE; 
    ELSIF ((x0 = FALSE) AND  (t0.Q = FALSE) AND  (t1.Q = TRUE)) THEN 
        cstate16 := 34932; y0 := FALSE; y1 := FALSE; y2 := FALSE; t0_start := FALSE;t1_start := FALSE; 
    ELSIF ((x0 = FALSE) AND  (t0.Q = TRUE) AND  (t1.Q = FALSE)) THEN 
        cstate16 := 28787; y0 := FALSE; y1 := FALSE; y2 := FALSE; t0_start := FALSE;t1_start := FALSE; 
    ELSIF ((x0 = FALSE) AND  (t0.Q = TRUE) AND  (t1.Q = TRUE)) THEN 
        cstate16 := 28788; y0 := FALSE; y1 := FALSE; y2 := FALSE; t0_start := FALSE;t1_start := FALSE; 
    ELSIF ((x0 = TRUE) AND  (t0.Q = FALSE) AND  (t1.Q = FALSE)) THEN 
        cstate16 := 48650; y0 := TRUE; y1 := TRUE; y2 := TRUE; t0_start := FALSE;t1_start := FALSE; 
    ELSIF ((x0 = TRUE) AND  (t0.Q = FALSE) AND  (t1.Q = TRUE)) THEN 
        cstate16 := 48646; y0 := TRUE; y1 := TRUE; y2 := TRUE; t0_start := FALSE;t1_start := FALSE; 
    ELSIF ((x0 = TRUE) AND  (t0.Q = TRUE) AND  (t1.Q = FALSE)) THEN 
        cstate16 := 43530; y0 := TRUE; y1 := TRUE; y2 := TRUE; t0_start := FALSE;t1_start := FALSE; 
    ELSIF ((x0 = TRUE) AND  (t0.Q = TRUE) AND  (t1.Q = TRUE)) THEN 
        cstate16 := 43526; y0 := TRUE; y1 := TRUE; y2 := TRUE; t0_start := FALSE;t1_start := FALSE; 
    END_IF;
48534:
    IF ((x0 = FALSE) AND  (t0.Q = FALSE) AND  (t1.Q = FALSE)) THEN 
        cstate16 := 34931; y0 := FALSE; y1 := FALSE; y2 := FALSE; t0_start := FALSE;t1_start := FALSE; 
    ELSIF ((x0 = FALSE) AND  (t0.Q = FALSE) AND  (t1.Q = TRUE)) THEN 
        cstate16 := 34932; y0 := FALSE; y1 := FALSE; y2 := FALSE; t0_start := FALSE;t1_start := FALSE; 
    ELSIF ((x0 = FALSE) AND  (t0.Q = TRUE) AND  (t1.Q = FALSE)) THEN 
        cstate16 := 27731; y0 := FALSE; y1 := FALSE; y2 := FALSE; t0_start := FALSE;t1_start := TRUE; t1_up := FALSE; 
    ELSIF ((x0 = FALSE) AND  (t0.Q = TRUE) AND  (t1.Q = TRUE)) THEN 
        cstate16 := 27732; y0 := FALSE; y1 := FALSE; y2 := FALSE; t0_start := FALSE;t1_start := TRUE; t1_up := FALSE; 
    ELSIF ((x0 = TRUE) AND  (t0.Q = FALSE) AND  (t1.Q = FALSE)) THEN 
        cstate16 := 48538; y0 := TRUE; y1 := FALSE; y2 := TRUE; t0_start := FALSE;t1_start := FALSE; 
    ELSIF ((x0 = TRUE) AND  (t0.Q = FALSE) AND  (t1.Q = TRUE)) THEN 
        cstate16 := 48534; y0 := TRUE; y1 := FALSE; y2 := TRUE; t0_start := FALSE;t1_start := FALSE; 
    ELSIF ((x0 = TRUE) AND  (t0.Q = TRUE) AND  (t1.Q = FALSE)) THEN 
        cstate16 := 42457; y0 := TRUE; y1 := TRUE; y2 := TRUE; t0_start := FALSE;t1_start := TRUE; t1_up := FALSE; 
    ELSIF ((x0 = TRUE) AND  (t0.Q = TRUE) AND  (t1.Q = TRUE)) THEN 
        cstate16 := 42453; y0 := TRUE; y1 := TRUE; y2 := TRUE; t0_start := FALSE;t1_start := TRUE; t1_up := FALSE; 
    END_IF;
0:
    IF ((x0 = FALSE) AND  (t0.Q = FALSE) AND  (t1.Q = FALSE)) THEN 
        cstate16 := 12353; y0 := FALSE; y1 := FALSE; y2 := FALSE; t0_start := FALSE;t1_start := FALSE; 
    ELSIF ((x0 = FALSE) AND  (t0.Q = FALSE) AND  (t1.Q = TRUE)) THEN 
        cstate16 := 12354; y0 := FALSE; y1 := FALSE; y2 := FALSE; t0_start := FALSE;t1_start := FALSE; 
    ELSIF ((x0 = FALSE) AND  (t0.Q = TRUE) AND  (t1.Q = FALSE)) THEN 
        cstate16 := 2113; y0 := FALSE; y1 := FALSE; y2 := FALSE; t0_start := FALSE;t1_start := FALSE; 
    ELSIF ((x0 = FALSE) AND  (t0.Q = TRUE) AND  (t1.Q = TRUE)) THEN 
        cstate16 := 2114; y0 := FALSE; y1 := FALSE; y2 := FALSE; t0_start := FALSE;t1_start := FALSE; 
    ELSIF ((x0 = TRUE) AND  (t0.Q = FALSE) AND  (t1.Q = FALSE)) THEN 
        cstate16 := 14401; y0 := FALSE; y1 := FALSE; y2 := FALSE; t0_start := FALSE;t1_start := FALSE; 
    ELSIF ((x0 = TRUE) AND  (t0.Q = FALSE) AND  (t1.Q = TRUE)) THEN 
        cstate16 := 14402; y0 := FALSE; y1 := FALSE; y2 := FALSE; t0_start := FALSE;t1_start := FALSE; 
    ELSIF ((x0 = TRUE) AND  (t0.Q = TRUE) AND  (t1.Q = FALSE)) THEN 
        cstate16 := 6209; y0 := FALSE; y1 := FALSE; y2 := FALSE; t0_start := FALSE;t1_start := FALSE; 
    ELSIF ((x0 = TRUE) AND  (t0.Q = TRUE) AND  (t1.Q = TRUE)) THEN 
        cstate16 := 6210; y0 := FALSE; y1 := FALSE; y2 := FALSE; t0_start := FALSE;t1_start := FALSE; 
    END_IF;
47692:
    IF ((x0 = FALSE) AND  (t0.Q = FALSE) AND  (t1.Q = FALSE)) THEN 
        cstate16 := 34931; y0 := FALSE; y1 := FALSE; y2 := FALSE; t0_start := FALSE;t1_start := FALSE; 
    ELSIF ((x0 = FALSE) AND  (t0.Q = FALSE) AND  (t1.Q = TRUE)) THEN 
        cstate16 := 34932; y0 := FALSE; y1 := FALSE; y2 := FALSE; t0_start := FALSE;t1_start := FALSE; 
    ELSIF ((x0 = FALSE) AND  (t0.Q = TRUE) AND  (t1.Q = FALSE)) THEN 
        cstate16 := 28787; y0 := FALSE; y1 := FALSE; y2 := FALSE; t0_start := FALSE;t1_start := FALSE; 
    ELSIF ((x0 = FALSE) AND  (t0.Q = TRUE) AND  (t1.Q = TRUE)) THEN 
        cstate16 := 28788; y0 := FALSE; y1 := FALSE; y2 := FALSE; t0_start := FALSE;t1_start := FALSE; 
    ELSIF ((x0 = TRUE) AND  (t0.Q = FALSE) AND  (t1.Q = FALSE)) THEN 
        cstate16 := 40172; y0 := TRUE; y1 := FALSE; y2 := TRUE; t0_start := TRUE; t0_up := FALSE;t1_start := FALSE; 
    ELSIF ((x0 = TRUE) AND  (t0.Q = FALSE) AND  (t1.Q = TRUE)) THEN 
        cstate16 := 40167; y0 := TRUE; y1 := FALSE; y2 := TRUE; t0_start := TRUE; t0_up := FALSE;t1_start := FALSE; 
    ELSIF ((x0 = TRUE) AND  (t0.Q = TRUE) AND  (t1.Q = FALSE)) THEN 
        cstate16 := 47692; y0 := TRUE; y1 := FALSE; y2 := TRUE; t0_start := FALSE;t1_start := FALSE; 
    ELSIF ((x0 = TRUE) AND  (t0.Q = TRUE) AND  (t1.Q = TRUE)) THEN 
        cstate16 := 47687; y0 := TRUE; y1 := FALSE; y2 := TRUE; t0_start := FALSE;t1_start := FALSE; 
    END_IF;
48538:
    IF ((x0 = FALSE) AND  (t0.Q = FALSE) AND  (t1.Q = FALSE)) THEN 
        cstate16 := 34931; y0 := FALSE; y1 := FALSE; y2 := FALSE; t0_start := FALSE;t1_start := FALSE; 
    ELSIF ((x0 = FALSE) AND  (t0.Q = FALSE) AND  (t1.Q = TRUE)) THEN 
        cstate16 := 34932; y0 := FALSE; y1 := FALSE; y2 := FALSE; t0_start := FALSE;t1_start := FALSE; 
    ELSIF ((x0 = FALSE) AND  (t0.Q = TRUE) AND  (t1.Q = FALSE)) THEN 
        cstate16 := 27731; y0 := FALSE; y1 := FALSE; y2 := FALSE; t0_start := FALSE;t1_start := TRUE; t1_up := FALSE; 
    ELSIF ((x0 = FALSE) AND  (t0.Q = TRUE) AND  (t1.Q = TRUE)) THEN 
        cstate16 := 27732; y0 := FALSE; y1 := FALSE; y2 := FALSE; t0_start := FALSE;t1_start := TRUE; t1_up := FALSE; 
    ELSIF ((x0 = TRUE) AND  (t0.Q = FALSE) AND  (t1.Q = FALSE)) THEN 
        cstate16 := 48538; y0 := TRUE; y1 := FALSE; y2 := TRUE; t0_start := FALSE;t1_start := FALSE; 
    ELSIF ((x0 = TRUE) AND  (t0.Q = FALSE) AND  (t1.Q = TRUE)) THEN 
        cstate16 := 48534; y0 := TRUE; y1 := FALSE; y2 := TRUE; t0_start := FALSE;t1_start := FALSE; 
    ELSIF ((x0 = TRUE) AND  (t0.Q = TRUE) AND  (t1.Q = FALSE)) THEN 
        cstate16 := 42457; y0 := TRUE; y1 := TRUE; y2 := TRUE; t0_start := FALSE;t1_start := TRUE; t1_up := FALSE; 
    ELSIF ((x0 = TRUE) AND  (t0.Q = TRUE) AND  (t1.Q = TRUE)) THEN 
        cstate16 := 42453; y0 := TRUE; y1 := TRUE; y2 := TRUE; t0_start := FALSE;t1_start := TRUE; t1_up := FALSE; 
    END_IF;
14401:
    IF ((x0 = FALSE) AND  (t0.Q = FALSE) AND  (t1.Q = FALSE)) THEN 
        cstate16 := 34931; y0 := FALSE; y1 := FALSE; y2 := FALSE; t0_start := FALSE;t1_start := FALSE; 
    ELSIF ((x0 = FALSE) AND  (t0.Q = FALSE) AND  (t1.Q = TRUE)) THEN 
        cstate16 := 34932; y0 := FALSE; y1 := FALSE; y2 := FALSE; t0_start := FALSE;t1_start := FALSE; 
    ELSIF ((x0 = FALSE) AND  (t0.Q = TRUE) AND  (t1.Q = FALSE)) THEN 
        cstate16 := 27731; y0 := FALSE; y1 := FALSE; y2 := FALSE; t0_start := FALSE;t1_start := TRUE; t1_up := FALSE; 
    ELSIF ((x0 = FALSE) AND  (t0.Q = TRUE) AND  (t1.Q = TRUE)) THEN 
        cstate16 := 27732; y0 := FALSE; y1 := FALSE; y2 := FALSE; t0_start := FALSE;t1_start := TRUE; t1_up := FALSE; 
    ELSIF ((x0 = TRUE) AND  (t0.Q = FALSE) AND  (t1.Q = FALSE)) THEN 
        cstate16 := 14401; y0 := FALSE; y1 := FALSE; y2 := FALSE; t0_start := FALSE;t1_start := FALSE; 
    ELSIF ((x0 = TRUE) AND  (t0.Q = FALSE) AND  (t1.Q = TRUE)) THEN 
        cstate16 := 14406; y0 := FALSE; y1 := FALSE; y2 := TRUE; t0_start := FALSE;t1_start := FALSE; 
    ELSIF ((x0 = TRUE) AND  (t0.Q = TRUE) AND  (t1.Q = FALSE)) THEN 
        cstate16 := 8353; y0 := FALSE; y1 := TRUE; y2 := FALSE; t0_start := FALSE;t1_start := TRUE; t1_up := FALSE; 
    ELSIF ((x0 = TRUE) AND  (t0.Q = TRUE) AND  (t1.Q = TRUE)) THEN 
        cstate16 := 8357; y0 := FALSE; y1 := TRUE; y2 := TRUE; t0_start := FALSE;t1_start := TRUE; t1_up := FALSE; 
    END_IF;
14402:
    IF ((x0 = FALSE) AND  (t0.Q = FALSE) AND  (t1.Q = FALSE)) THEN 
        cstate16 := 34931; y0 := FALSE; y1 := FALSE; y2 := FALSE; t0_start := FALSE;t1_start := FALSE; 
    ELSIF ((x0 = FALSE) AND  (t0.Q = FALSE) AND  (t1.Q = TRUE)) THEN 
        cstate16 := 34932; y0 := FALSE; y1 := FALSE; y2 := FALSE; t0_start := FALSE;t1_start := FALSE; 
    ELSIF ((x0 = FALSE) AND  (t0.Q = TRUE) AND  (t1.Q = FALSE)) THEN 
        cstate16 := 27731; y0 := FALSE; y1 := FALSE; y2 := FALSE; t0_start := FALSE;t1_start := TRUE; t1_up := FALSE; 
    ELSIF ((x0 = FALSE) AND  (t0.Q = TRUE) AND  (t1.Q = TRUE)) THEN 
        cstate16 := 27732; y0 := FALSE; y1 := FALSE; y2 := FALSE; t0_start := FALSE;t1_start := TRUE; t1_up := FALSE; 
    ELSIF ((x0 = TRUE) AND  (t0.Q = FALSE) AND  (t1.Q = FALSE)) THEN 
        cstate16 := 14401; y0 := FALSE; y1 := FALSE; y2 := FALSE; t0_start := FALSE;t1_start := FALSE; 
    ELSIF ((x0 = TRUE) AND  (t0.Q = FALSE) AND  (t1.Q = TRUE)) THEN 
        cstate16 := 14402; y0 := FALSE; y1 := FALSE; y2 := FALSE; t0_start := FALSE;t1_start := FALSE; 
    ELSIF ((x0 = TRUE) AND  (t0.Q = TRUE) AND  (t1.Q = FALSE)) THEN 
        cstate16 := 8353; y0 := FALSE; y1 := TRUE; y2 := FALSE; t0_start := FALSE;t1_start := TRUE; t1_up := FALSE; 
    ELSIF ((x0 = TRUE) AND  (t0.Q = TRUE) AND  (t1.Q = TRUE)) THEN 
        cstate16 := 8354; y0 := FALSE; y1 := TRUE; y2 := FALSE; t0_start := FALSE;t1_start := TRUE; t1_up := FALSE; 
    END_IF;
38148:
    IF ((x0 = FALSE) AND  (t0.Q = FALSE) AND  (t1.Q = FALSE)) THEN 
        cstate16 := 23667; y0 := FALSE; y1 := FALSE; y2 := FALSE; t0_start := FALSE;t1_start := FALSE; 
    ELSIF ((x0 = FALSE) AND  (t0.Q = FALSE) AND  (t1.Q = TRUE)) THEN 
        cstate16 := 26740; y0 := FALSE; y1 := FALSE; y2 := FALSE; t0_start := FALSE;t1_start := FALSE; 
    ELSIF ((x0 = FALSE) AND  (t0.Q = TRUE) AND  (t1.Q = FALSE)) THEN 
        cstate16 := 17523; y0 := FALSE; y1 := FALSE; y2 := FALSE; t0_start := FALSE;t1_start := FALSE; 
    ELSIF ((x0 = FALSE) AND  (t0.Q = TRUE) AND  (t1.Q = TRUE)) THEN 
        cstate16 := 22644; y0 := FALSE; y1 := FALSE; y2 := FALSE; t0_start := FALSE;t1_start := FALSE; 
    ELSIF ((x0 = TRUE) AND  (t0.Q = FALSE) AND  (t1.Q = FALSE)) THEN 
        cstate16 := 41699; y0 := TRUE; y1 := TRUE; y2 := FALSE; t0_start := FALSE;t1_start := FALSE; 
    ELSIF ((x0 = TRUE) AND  (t0.Q = FALSE) AND  (t1.Q = TRUE)) THEN 
        cstate16 := 40660; y0 := TRUE; y1 := TRUE; y2 := FALSE; t0_start := FALSE;t1_start := FALSE; 
    ELSIF ((x0 = TRUE) AND  (t0.Q = TRUE) AND  (t1.Q = FALSE)) THEN 
        cstate16 := 46739; y0 := TRUE; y1 := TRUE; y2 := FALSE; t0_start := FALSE;t1_start := FALSE; 
    ELSIF ((x0 = TRUE) AND  (t0.Q = TRUE) AND  (t1.Q = TRUE)) THEN 
        cstate16 := 47796; y0 := TRUE; y1 := TRUE; y2 := FALSE; t0_start := FALSE;t1_start := FALSE; 
    END_IF;
43522:
    IF ((x0 = FALSE) AND  (t0.Q = FALSE) AND  (t1.Q = FALSE)) THEN 
        cstate16 := 34931; y0 := FALSE; y1 := FALSE; y2 := FALSE; t0_start := FALSE;t1_start := FALSE; 
    ELSIF ((x0 = FALSE) AND  (t0.Q = FALSE) AND  (t1.Q = TRUE)) THEN 
        cstate16 := 34932; y0 := FALSE; y1 := FALSE; y2 := FALSE; t0_start := FALSE;t1_start := FALSE; 
    ELSIF ((x0 = FALSE) AND  (t0.Q = TRUE) AND  (t1.Q = FALSE)) THEN 
        cstate16 := 28787; y0 := FALSE; y1 := FALSE; y2 := FALSE; t0_start := FALSE;t1_start := FALSE; 
    ELSIF ((x0 = FALSE) AND  (t0.Q = TRUE) AND  (t1.Q = TRUE)) THEN 
        cstate16 := 28788; y0 := FALSE; y1 := FALSE; y2 := FALSE; t0_start := FALSE;t1_start := FALSE; 
    ELSIF ((x0 = TRUE) AND  (t0.Q = FALSE) AND  (t1.Q = FALSE)) THEN 
        cstate16 := 48641; y0 := TRUE; y1 := TRUE; y2 := FALSE; t0_start := FALSE;t1_start := FALSE; 
    ELSIF ((x0 = TRUE) AND  (t0.Q = FALSE) AND  (t1.Q = TRUE)) THEN 
        cstate16 := 48642; y0 := TRUE; y1 := TRUE; y2 := FALSE; t0_start := FALSE;t1_start := FALSE; 
    ELSIF ((x0 = TRUE) AND  (t0.Q = TRUE) AND  (t1.Q = FALSE)) THEN 
        cstate16 := 43521; y0 := TRUE; y1 := TRUE; y2 := FALSE; t0_start := FALSE;t1_start := FALSE; 
    ELSIF ((x0 = TRUE) AND  (t0.Q = TRUE) AND  (t1.Q = TRUE)) THEN 
        cstate16 := 43522; y0 := TRUE; y1 := TRUE; y2 := FALSE; t0_start := FALSE;t1_start := FALSE; 
    END_IF;
14673:
    IF ((x0 = FALSE) AND  (t0.Q = FALSE) AND  (t1.Q = FALSE)) THEN 
        cstate16 := 34931; y0 := FALSE; y1 := FALSE; y2 := FALSE; t0_start := FALSE;t1_start := FALSE; 
    ELSIF ((x0 = FALSE) AND  (t0.Q = FALSE) AND  (t1.Q = TRUE)) THEN 
        cstate16 := 34932; y0 := FALSE; y1 := FALSE; y2 := FALSE; t0_start := FALSE;t1_start := FALSE; 
    ELSIF ((x0 = FALSE) AND  (t0.Q = TRUE) AND  (t1.Q = FALSE)) THEN 
        cstate16 := 27731; y0 := FALSE; y1 := FALSE; y2 := FALSE; t0_start := FALSE;t1_start := TRUE; t1_up := FALSE; 
    ELSIF ((x0 = FALSE) AND  (t0.Q = TRUE) AND  (t1.Q = TRUE)) THEN 
        cstate16 := 27732; y0 := FALSE; y1 := FALSE; y2 := FALSE; t0_start := FALSE;t1_start := TRUE; t1_up := FALSE; 
    ELSIF ((x0 = TRUE) AND  (t0.Q = FALSE) AND  (t1.Q = FALSE)) THEN 
        cstate16 := 14673; y0 := FALSE; y1 := TRUE; y2 := FALSE; t0_start := FALSE;t1_start := FALSE; 
    ELSIF ((x0 = TRUE) AND  (t0.Q = FALSE) AND  (t1.Q = TRUE)) THEN 
        cstate16 := 14678; y0 := FALSE; y1 := TRUE; y2 := TRUE; t0_start := FALSE;t1_start := FALSE; 
    ELSIF ((x0 = TRUE) AND  (t0.Q = TRUE) AND  (t1.Q = FALSE)) THEN 
        cstate16 := 8353; y0 := FALSE; y1 := TRUE; y2 := FALSE; t0_start := FALSE;t1_start := TRUE; t1_up := FALSE; 
    ELSIF ((x0 = TRUE) AND  (t0.Q = TRUE) AND  (t1.Q = TRUE)) THEN 
        cstate16 := 8357; y0 := FALSE; y1 := TRUE; y2 := TRUE; t0_start := FALSE;t1_start := TRUE; t1_up := FALSE; 
    END_IF;
25121:
    IF ((x0 = FALSE) AND  (t0.Q = FALSE) AND  (t1.Q = FALSE)) THEN 
        cstate16 := 23667; y0 := FALSE; y1 := FALSE; y2 := FALSE; t0_start := FALSE;t1_start := FALSE; 
    ELSIF ((x0 = FALSE) AND  (t0.Q = FALSE) AND  (t1.Q = TRUE)) THEN 
        cstate16 := 26740; y0 := FALSE; y1 := FALSE; y2 := FALSE; t0_start := FALSE;t1_start := FALSE; 
    ELSIF ((x0 = FALSE) AND  (t0.Q = TRUE) AND  (t1.Q = FALSE)) THEN 
        cstate16 := 17491; y0 := FALSE; y1 := FALSE; y2 := FALSE; t0_start := FALSE;t1_start := TRUE; t1_up := FALSE; 
    ELSIF ((x0 = FALSE) AND  (t0.Q = TRUE) AND  (t1.Q = TRUE)) THEN 
        cstate16 := 17492; y0 := FALSE; y1 := FALSE; y2 := FALSE; t0_start := FALSE;t1_start := TRUE; t1_up := FALSE; 
    ELSIF ((x0 = TRUE) AND  (t0.Q = FALSE) AND  (t1.Q = FALSE)) THEN 
        cstate16 := 25121; y0 := TRUE; y1 := TRUE; y2 := FALSE; t0_start := FALSE;t1_start := FALSE; 
    ELSIF ((x0 = TRUE) AND  (t0.Q = FALSE) AND  (t1.Q = TRUE)) THEN 
        cstate16 := 26134; y0 := TRUE; y1 := TRUE; y2 := TRUE; t0_start := FALSE;t1_start := FALSE; 
    ELSIF ((x0 = TRUE) AND  (t0.Q = TRUE) AND  (t1.Q = FALSE)) THEN 
        cstate16 := 42449; y0 := TRUE; y1 := TRUE; y2 := FALSE; t0_start := FALSE;t1_start := TRUE; t1_up := FALSE; 
    ELSIF ((x0 = TRUE) AND  (t0.Q = TRUE) AND  (t1.Q = TRUE)) THEN 
        cstate16 := 42453; y0 := TRUE; y1 := TRUE; y2 := TRUE; t0_start := FALSE;t1_start := TRUE; t1_up := FALSE; 
    END_IF;
43521:
    IF ((x0 = FALSE) AND  (t0.Q = FALSE) AND  (t1.Q = FALSE)) THEN 
        cstate16 := 34931; y0 := FALSE; y1 := FALSE; y2 := FALSE; t0_start := FALSE;t1_start := FALSE; 
    ELSIF ((x0 = FALSE) AND  (t0.Q = FALSE) AND  (t1.Q = TRUE)) THEN 
        cstate16 := 34932; y0 := FALSE; y1 := FALSE; y2 := FALSE; t0_start := FALSE;t1_start := FALSE; 
    ELSIF ((x0 = FALSE) AND  (t0.Q = TRUE) AND  (t1.Q = FALSE)) THEN 
        cstate16 := 28787; y0 := FALSE; y1 := FALSE; y2 := FALSE; t0_start := FALSE;t1_start := FALSE; 
    ELSIF ((x0 = FALSE) AND  (t0.Q = TRUE) AND  (t1.Q = TRUE)) THEN 
        cstate16 := 28788; y0 := FALSE; y1 := FALSE; y2 := FALSE; t0_start := FALSE;t1_start := FALSE; 
    ELSIF ((x0 = TRUE) AND  (t0.Q = FALSE) AND  (t1.Q = FALSE)) THEN 
        cstate16 := 48641; y0 := TRUE; y1 := TRUE; y2 := FALSE; t0_start := FALSE;t1_start := FALSE; 
    ELSIF ((x0 = TRUE) AND  (t0.Q = FALSE) AND  (t1.Q = TRUE)) THEN 
        cstate16 := 48646; y0 := TRUE; y1 := TRUE; y2 := TRUE; t0_start := FALSE;t1_start := FALSE; 
    ELSIF ((x0 = TRUE) AND  (t0.Q = TRUE) AND  (t1.Q = FALSE)) THEN 
        cstate16 := 43521; y0 := TRUE; y1 := TRUE; y2 := FALSE; t0_start := FALSE;t1_start := FALSE; 
    ELSIF ((x0 = TRUE) AND  (t0.Q = TRUE) AND  (t1.Q = TRUE)) THEN 
        cstate16 := 43526; y0 := TRUE; y1 := TRUE; y2 := TRUE; t0_start := FALSE;t1_start := FALSE; 
    END_IF;
14406:
    IF ((x0 = FALSE) AND  (t0.Q = FALSE) AND  (t1.Q = FALSE)) THEN 
        cstate16 := 34931; y0 := FALSE; y1 := FALSE; y2 := FALSE; t0_start := FALSE;t1_start := FALSE; 
    ELSIF ((x0 = FALSE) AND  (t0.Q = FALSE) AND  (t1.Q = TRUE)) THEN 
        cstate16 := 34932; y0 := FALSE; y1 := FALSE; y2 := FALSE; t0_start := FALSE;t1_start := FALSE; 
    ELSIF ((x0 = FALSE) AND  (t0.Q = TRUE) AND  (t1.Q = FALSE)) THEN 
        cstate16 := 27731; y0 := FALSE; y1 := FALSE; y2 := FALSE; t0_start := FALSE;t1_start := TRUE; t1_up := FALSE; 
    ELSIF ((x0 = FALSE) AND  (t0.Q = TRUE) AND  (t1.Q = TRUE)) THEN 
        cstate16 := 27732; y0 := FALSE; y1 := FALSE; y2 := FALSE; t0_start := FALSE;t1_start := TRUE; t1_up := FALSE; 
    ELSIF ((x0 = TRUE) AND  (t0.Q = FALSE) AND  (t1.Q = FALSE)) THEN 
        cstate16 := 14410; y0 := FALSE; y1 := FALSE; y2 := TRUE; t0_start := FALSE;t1_start := FALSE; 
    ELSIF ((x0 = TRUE) AND  (t0.Q = FALSE) AND  (t1.Q = TRUE)) THEN 
        cstate16 := 14406; y0 := FALSE; y1 := FALSE; y2 := TRUE; t0_start := FALSE;t1_start := FALSE; 
    ELSIF ((x0 = TRUE) AND  (t0.Q = TRUE) AND  (t1.Q = FALSE)) THEN 
        cstate16 := 8361; y0 := FALSE; y1 := TRUE; y2 := TRUE; t0_start := FALSE;t1_start := TRUE; t1_up := FALSE; 
    ELSIF ((x0 = TRUE) AND  (t0.Q = TRUE) AND  (t1.Q = TRUE)) THEN 
        cstate16 := 8357; y0 := FALSE; y1 := TRUE; y2 := TRUE; t0_start := FALSE;t1_start := TRUE; t1_up := FALSE; 
    END_IF;
49657:
    IF ((x0 = FALSE) AND  (t0.Q = FALSE) AND  (t1.Q = FALSE)) THEN 
        cstate16 := 32883; y0 := FALSE; y1 := FALSE; y2 := FALSE; t0_start := FALSE;t1_start := FALSE; 
    ELSIF ((x0 = FALSE) AND  (t0.Q = FALSE) AND  (t1.Q = TRUE)) THEN 
        cstate16 := 34932; y0 := FALSE; y1 := FALSE; y2 := FALSE; t0_start := FALSE;t1_start := FALSE; 
    ELSIF ((x0 = FALSE) AND  (t0.Q = TRUE) AND  (t1.Q = FALSE)) THEN 
        cstate16 := 27731; y0 := FALSE; y1 := FALSE; y2 := FALSE; t0_start := FALSE;t1_start := TRUE; t1_up := FALSE; 
    ELSIF ((x0 = FALSE) AND  (t0.Q = TRUE) AND  (t1.Q = TRUE)) THEN 
        cstate16 := 27732; y0 := FALSE; y1 := FALSE; y2 := FALSE; t0_start := FALSE;t1_start := TRUE; t1_up := FALSE; 
    ELSIF ((x0 = TRUE) AND  (t0.Q = FALSE) AND  (t1.Q = FALSE)) THEN 
        cstate16 := 49657; y0 := TRUE; y1 := TRUE; y2 := TRUE; t0_start := FALSE;t1_start := FALSE; 
    ELSIF ((x0 = TRUE) AND  (t0.Q = FALSE) AND  (t1.Q = TRUE)) THEN 
        cstate16 := 48646; y0 := TRUE; y1 := TRUE; y2 := TRUE; t0_start := FALSE;t1_start := FALSE; 
    ELSIF ((x0 = TRUE) AND  (t0.Q = TRUE) AND  (t1.Q = FALSE)) THEN 
        cstate16 := 42457; y0 := TRUE; y1 := TRUE; y2 := TRUE; t0_start := FALSE;t1_start := TRUE; t1_up := FALSE; 
    ELSIF ((x0 = TRUE) AND  (t0.Q = TRUE) AND  (t1.Q = TRUE)) THEN 
        cstate16 := 42453; y0 := TRUE; y1 := TRUE; y2 := TRUE; t0_start := FALSE;t1_start := TRUE; t1_up := FALSE; 
    END_IF;
41643:
    IF ((x0 = FALSE) AND  (t0.Q = FALSE) AND  (t1.Q = FALSE)) THEN 
        cstate16 := 23667; y0 := FALSE; y1 := FALSE; y2 := FALSE; t0_start := FALSE;t1_start := FALSE; 
    ELSIF ((x0 = FALSE) AND  (t0.Q = FALSE) AND  (t1.Q = TRUE)) THEN 
        cstate16 := 26740; y0 := FALSE; y1 := FALSE; y2 := FALSE; t0_start := FALSE;t1_start := FALSE; 
    ELSIF ((x0 = FALSE) AND  (t0.Q = TRUE) AND  (t1.Q = FALSE)) THEN 
        cstate16 := 17491; y0 := FALSE; y1 := FALSE; y2 := FALSE; t0_start := FALSE;t1_start := TRUE; t1_up := FALSE; 
    ELSIF ((x0 = FALSE) AND  (t0.Q = TRUE) AND  (t1.Q = TRUE)) THEN 
        cstate16 := 17492; y0 := FALSE; y1 := FALSE; y2 := FALSE; t0_start := FALSE;t1_start := TRUE; t1_up := FALSE; 
    ELSIF ((x0 = TRUE) AND  (t0.Q = FALSE) AND  (t1.Q = FALSE)) THEN 
        cstate16 := 41707; y0 := TRUE; y1 := TRUE; y2 := TRUE; t0_start := FALSE;t1_start := FALSE; 
    ELSIF ((x0 = TRUE) AND  (t0.Q = FALSE) AND  (t1.Q = TRUE)) THEN 
        cstate16 := 40663; y0 := TRUE; y1 := TRUE; y2 := TRUE; t0_start := FALSE;t1_start := FALSE; 
    ELSIF ((x0 = TRUE) AND  (t0.Q = TRUE) AND  (t1.Q = FALSE)) THEN 
        cstate16 := 46651; y0 := TRUE; y1 := TRUE; y2 := TRUE; t0_start := FALSE;t1_start := TRUE; t1_up := FALSE; 
    ELSIF ((x0 = TRUE) AND  (t0.Q = TRUE) AND  (t1.Q = TRUE)) THEN 
        cstate16 := 46648; y0 := TRUE; y1 := TRUE; y2 := TRUE; t0_start := FALSE;t1_start := TRUE; t1_up := FALSE; 
    END_IF;
12353:
    IF ((x0 = FALSE) AND  (t0.Q = FALSE) AND  (t1.Q = FALSE)) THEN 
        cstate16 := 34931; y0 := FALSE; y1 := FALSE; y2 := FALSE; t0_start := FALSE;t1_start := FALSE; 
    ELSIF ((x0 = FALSE) AND  (t0.Q = FALSE) AND  (t1.Q = TRUE)) THEN 
        cstate16 := 34932; y0 := FALSE; y1 := FALSE; y2 := FALSE; t0_start := FALSE;t1_start := FALSE; 
    ELSIF ((x0 = FALSE) AND  (t0.Q = TRUE) AND  (t1.Q = FALSE)) THEN 
        cstate16 := 27731; y0 := FALSE; y1 := FALSE; y2 := FALSE; t0_start := FALSE;t1_start := TRUE; t1_up := FALSE; 
    ELSIF ((x0 = FALSE) AND  (t0.Q = TRUE) AND  (t1.Q = TRUE)) THEN 
        cstate16 := 27732; y0 := FALSE; y1 := FALSE; y2 := FALSE; t0_start := FALSE;t1_start := TRUE; t1_up := FALSE; 
    ELSIF ((x0 = TRUE) AND  (t0.Q = FALSE) AND  (t1.Q = FALSE)) THEN 
        cstate16 := 25793; y0 := TRUE; y1 := FALSE; y2 := FALSE; t0_start := TRUE; t0_up := FALSE;t1_start := FALSE; 
    ELSIF ((x0 = TRUE) AND  (t0.Q = FALSE) AND  (t1.Q = TRUE)) THEN 
        cstate16 := 25798; y0 := TRUE; y1 := FALSE; y2 := TRUE; t0_start := TRUE; t0_up := FALSE;t1_start := FALSE; 
    ELSIF ((x0 = TRUE) AND  (t0.Q = TRUE) AND  (t1.Q = FALSE)) THEN 
        cstate16 := 19665; y0 := TRUE; y1 := TRUE; y2 := FALSE; t0_start := TRUE; t0_up := FALSE;t1_start := TRUE; t1_up := FALSE; 
    ELSIF ((x0 = TRUE) AND  (t0.Q = TRUE) AND  (t1.Q = TRUE)) THEN 
        cstate16 := 19669; y0 := TRUE; y1 := TRUE; y2 := TRUE; t0_start := TRUE; t0_up := FALSE;t1_start := TRUE; t1_up := FALSE; 
    END_IF;
12354:
    IF ((x0 = FALSE) AND  (t0.Q = FALSE) AND  (t1.Q = FALSE)) THEN 
        cstate16 := 34931; y0 := FALSE; y1 := FALSE; y2 := FALSE; t0_start := FALSE;t1_start := FALSE; 
    ELSIF ((x0 = FALSE) AND  (t0.Q = FALSE) AND  (t1.Q = TRUE)) THEN 
        cstate16 := 34932; y0 := FALSE; y1 := FALSE; y2 := FALSE; t0_start := FALSE;t1_start := FALSE; 
    ELSIF ((x0 = FALSE) AND  (t0.Q = TRUE) AND  (t1.Q = FALSE)) THEN 
        cstate16 := 27731; y0 := FALSE; y1 := FALSE; y2 := FALSE; t0_start := FALSE;t1_start := TRUE; t1_up := FALSE; 
    ELSIF ((x0 = FALSE) AND  (t0.Q = TRUE) AND  (t1.Q = TRUE)) THEN 
        cstate16 := 27732; y0 := FALSE; y1 := FALSE; y2 := FALSE; t0_start := FALSE;t1_start := TRUE; t1_up := FALSE; 
    ELSIF ((x0 = TRUE) AND  (t0.Q = FALSE) AND  (t1.Q = FALSE)) THEN 
        cstate16 := 25793; y0 := TRUE; y1 := FALSE; y2 := FALSE; t0_start := TRUE; t0_up := FALSE;t1_start := FALSE; 
    ELSIF ((x0 = TRUE) AND  (t0.Q = FALSE) AND  (t1.Q = TRUE)) THEN 
        cstate16 := 25794; y0 := TRUE; y1 := FALSE; y2 := FALSE; t0_start := TRUE; t0_up := FALSE;t1_start := FALSE; 
    ELSIF ((x0 = TRUE) AND  (t0.Q = TRUE) AND  (t1.Q = FALSE)) THEN 
        cstate16 := 19665; y0 := TRUE; y1 := TRUE; y2 := FALSE; t0_start := TRUE; t0_up := FALSE;t1_start := TRUE; t1_up := FALSE; 
    ELSIF ((x0 = TRUE) AND  (t0.Q = TRUE) AND  (t1.Q = TRUE)) THEN 
        cstate16 := 19666; y0 := TRUE; y1 := TRUE; y2 := FALSE; t0_start := TRUE; t0_up := FALSE;t1_start := TRUE; t1_up := FALSE; 
    END_IF;
26739:
    IF ((x0 = FALSE) AND  (t0.Q = FALSE) AND  (t1.Q = FALSE)) THEN 
        cstate16 := 26739; y0 := FALSE; y1 := FALSE; y2 := FALSE; t0_start := FALSE;t1_start := FALSE; 
    ELSIF ((x0 = FALSE) AND  (t0.Q = FALSE) AND  (t1.Q = TRUE)) THEN 
        cstate16 := 26740; y0 := FALSE; y1 := FALSE; y2 := FALSE; t0_start := FALSE;t1_start := FALSE; 
    ELSIF ((x0 = FALSE) AND  (t0.Q = TRUE) AND  (t1.Q = FALSE)) THEN 
        cstate16 := 17491; y0 := FALSE; y1 := FALSE; y2 := FALSE; t0_start := FALSE;t1_start := TRUE; t1_up := FALSE; 
    ELSIF ((x0 = FALSE) AND  (t0.Q = TRUE) AND  (t1.Q = TRUE)) THEN 
        cstate16 := 17492; y0 := FALSE; y1 := FALSE; y2 := FALSE; t0_start := FALSE;t1_start := TRUE; t1_up := FALSE; 
    ELSIF ((x0 = TRUE) AND  (t0.Q = FALSE) AND  (t1.Q = FALSE)) THEN 
        cstate16 := 40163; y0 := TRUE; y1 := FALSE; y2 := FALSE; t0_start := TRUE; t0_up := FALSE;t1_start := FALSE; 
    ELSIF ((x0 = TRUE) AND  (t0.Q = FALSE) AND  (t1.Q = TRUE)) THEN 
        cstate16 := 40167; y0 := TRUE; y1 := FALSE; y2 := TRUE; t0_start := TRUE; t0_up := FALSE;t1_start := FALSE; 
    ELSIF ((x0 = TRUE) AND  (t0.Q = TRUE) AND  (t1.Q = FALSE)) THEN 
        cstate16 := 38147; y0 := TRUE; y1 := TRUE; y2 := FALSE; t0_start := TRUE; t0_up := FALSE;t1_start := TRUE; t1_up := FALSE; 
    ELSIF ((x0 = TRUE) AND  (t0.Q = TRUE) AND  (t1.Q = TRUE)) THEN 
        cstate16 := 38152; y0 := TRUE; y1 := TRUE; y2 := TRUE; t0_start := TRUE; t0_up := FALSE;t1_start := TRUE; t1_up := FALSE; 
    END_IF;
38115:
    IF ((x0 = FALSE) AND  (t0.Q = FALSE) AND  (t1.Q = FALSE)) THEN 
        cstate16 := 23667; y0 := FALSE; y1 := FALSE; y2 := FALSE; t0_start := FALSE;t1_start := FALSE; 
    ELSIF ((x0 = FALSE) AND  (t0.Q = FALSE) AND  (t1.Q = TRUE)) THEN 
        cstate16 := 26740; y0 := FALSE; y1 := FALSE; y2 := FALSE; t0_start := FALSE;t1_start := FALSE; 
    ELSIF ((x0 = FALSE) AND  (t0.Q = TRUE) AND  (t1.Q = FALSE)) THEN 
        cstate16 := 17523; y0 := FALSE; y1 := FALSE; y2 := FALSE; t0_start := FALSE;t1_start := FALSE; 
    ELSIF ((x0 = FALSE) AND  (t0.Q = TRUE) AND  (t1.Q = TRUE)) THEN 
        cstate16 := 22644; y0 := FALSE; y1 := FALSE; y2 := FALSE; t0_start := FALSE;t1_start := FALSE; 
    ELSIF ((x0 = TRUE) AND  (t0.Q = FALSE) AND  (t1.Q = FALSE)) THEN 
        cstate16 := 41555; y0 := TRUE; y1 := FALSE; y2 := FALSE; t0_start := FALSE;t1_start := FALSE; 
    ELSIF ((x0 = TRUE) AND  (t0.Q = FALSE) AND  (t1.Q = TRUE)) THEN 
        cstate16 := 40535; y0 := TRUE; y1 := FALSE; y2 := TRUE; t0_start := FALSE;t1_start := FALSE; 
    ELSIF ((x0 = TRUE) AND  (t0.Q = TRUE) AND  (t1.Q = FALSE)) THEN 
        cstate16 := 46659; y0 := TRUE; y1 := FALSE; y2 := FALSE; t0_start := FALSE;t1_start := FALSE; 
    ELSIF ((x0 = TRUE) AND  (t0.Q = TRUE) AND  (t1.Q = TRUE)) THEN 
        cstate16 := 47687; y0 := TRUE; y1 := FALSE; y2 := TRUE; t0_start := FALSE;t1_start := FALSE; 
    END_IF;
14410:
    IF ((x0 = FALSE) AND  (t0.Q = FALSE) AND  (t1.Q = FALSE)) THEN 
        cstate16 := 34931; y0 := FALSE; y1 := FALSE; y2 := FALSE; t0_start := FALSE;t1_start := FALSE; 
    ELSIF ((x0 = FALSE) AND  (t0.Q = FALSE) AND  (t1.Q = TRUE)) THEN 
        cstate16 := 34932; y0 := FALSE; y1 := FALSE; y2 := FALSE; t0_start := FALSE;t1_start := FALSE; 
    ELSIF ((x0 = FALSE) AND  (t0.Q = TRUE) AND  (t1.Q = FALSE)) THEN 
        cstate16 := 27731; y0 := FALSE; y1 := FALSE; y2 := FALSE; t0_start := FALSE;t1_start := TRUE; t1_up := FALSE; 
    ELSIF ((x0 = FALSE) AND  (t0.Q = TRUE) AND  (t1.Q = TRUE)) THEN 
        cstate16 := 27732; y0 := FALSE; y1 := FALSE; y2 := FALSE; t0_start := FALSE;t1_start := TRUE; t1_up := FALSE; 
    ELSIF ((x0 = TRUE) AND  (t0.Q = FALSE) AND  (t1.Q = FALSE)) THEN 
        cstate16 := 14410; y0 := FALSE; y1 := FALSE; y2 := TRUE; t0_start := FALSE;t1_start := FALSE; 
    ELSIF ((x0 = TRUE) AND  (t0.Q = FALSE) AND  (t1.Q = TRUE)) THEN 
        cstate16 := 14406; y0 := FALSE; y1 := FALSE; y2 := TRUE; t0_start := FALSE;t1_start := FALSE; 
    ELSIF ((x0 = TRUE) AND  (t0.Q = TRUE) AND  (t1.Q = FALSE)) THEN 
        cstate16 := 8361; y0 := FALSE; y1 := TRUE; y2 := TRUE; t0_start := FALSE;t1_start := TRUE; t1_up := FALSE; 
    ELSIF ((x0 = TRUE) AND  (t0.Q = TRUE) AND  (t1.Q = TRUE)) THEN 
        cstate16 := 8357; y0 := FALSE; y1 := TRUE; y2 := TRUE; t0_start := FALSE;t1_start := TRUE; t1_up := FALSE; 
    END_IF;
40540:
    IF ((x0 = FALSE) AND  (t0.Q = FALSE) AND  (t1.Q = FALSE)) THEN 
        cstate16 := 26739; y0 := FALSE; y1 := FALSE; y2 := FALSE; t0_start := FALSE;t1_start := FALSE; 
    ELSIF ((x0 = FALSE) AND  (t0.Q = FALSE) AND  (t1.Q = TRUE)) THEN 
        cstate16 := 26740; y0 := FALSE; y1 := FALSE; y2 := FALSE; t0_start := FALSE;t1_start := FALSE; 
    ELSIF ((x0 = FALSE) AND  (t0.Q = TRUE) AND  (t1.Q = FALSE)) THEN 
        cstate16 := 17491; y0 := FALSE; y1 := FALSE; y2 := FALSE; t0_start := FALSE;t1_start := TRUE; t1_up := FALSE; 
    ELSIF ((x0 = FALSE) AND  (t0.Q = TRUE) AND  (t1.Q = TRUE)) THEN 
        cstate16 := 17492; y0 := FALSE; y1 := FALSE; y2 := FALSE; t0_start := FALSE;t1_start := TRUE; t1_up := FALSE; 
    ELSIF ((x0 = TRUE) AND  (t0.Q = FALSE) AND  (t1.Q = FALSE)) THEN 
        cstate16 := 40540; y0 := TRUE; y1 := FALSE; y2 := TRUE; t0_start := FALSE;t1_start := FALSE; 
    ELSIF ((x0 = TRUE) AND  (t0.Q = FALSE) AND  (t1.Q = TRUE)) THEN 
        cstate16 := 40535; y0 := TRUE; y1 := FALSE; y2 := TRUE; t0_start := FALSE;t1_start := FALSE; 
    ELSIF ((x0 = TRUE) AND  (t0.Q = TRUE) AND  (t1.Q = FALSE)) THEN 
        cstate16 := 46651; y0 := TRUE; y1 := TRUE; y2 := TRUE; t0_start := FALSE;t1_start := TRUE; t1_up := FALSE; 
    ELSIF ((x0 = TRUE) AND  (t0.Q = TRUE) AND  (t1.Q = TRUE)) THEN 
        cstate16 := 46648; y0 := TRUE; y1 := TRUE; y2 := TRUE; t0_start := FALSE;t1_start := TRUE; t1_up := FALSE; 
    END_IF;
48529:
    IF ((x0 = FALSE) AND  (t0.Q = FALSE) AND  (t1.Q = FALSE)) THEN 
        cstate16 := 34931; y0 := FALSE; y1 := FALSE; y2 := FALSE; t0_start := FALSE;t1_start := FALSE; 
    ELSIF ((x0 = FALSE) AND  (t0.Q = FALSE) AND  (t1.Q = TRUE)) THEN 
        cstate16 := 34932; y0 := FALSE; y1 := FALSE; y2 := FALSE; t0_start := FALSE;t1_start := FALSE; 
    ELSIF ((x0 = FALSE) AND  (t0.Q = TRUE) AND  (t1.Q = FALSE)) THEN 
        cstate16 := 27731; y0 := FALSE; y1 := FALSE; y2 := FALSE; t0_start := FALSE;t1_start := TRUE; t1_up := FALSE; 
    ELSIF ((x0 = FALSE) AND  (t0.Q = TRUE) AND  (t1.Q = TRUE)) THEN 
        cstate16 := 27732; y0 := FALSE; y1 := FALSE; y2 := FALSE; t0_start := FALSE;t1_start := TRUE; t1_up := FALSE; 
    ELSIF ((x0 = TRUE) AND  (t0.Q = FALSE) AND  (t1.Q = FALSE)) THEN 
        cstate16 := 48529; y0 := TRUE; y1 := FALSE; y2 := FALSE; t0_start := FALSE;t1_start := FALSE; 
    ELSIF ((x0 = TRUE) AND  (t0.Q = FALSE) AND  (t1.Q = TRUE)) THEN 
        cstate16 := 48534; y0 := TRUE; y1 := FALSE; y2 := TRUE; t0_start := FALSE;t1_start := FALSE; 
    ELSIF ((x0 = TRUE) AND  (t0.Q = TRUE) AND  (t1.Q = FALSE)) THEN 
        cstate16 := 42449; y0 := TRUE; y1 := TRUE; y2 := FALSE; t0_start := FALSE;t1_start := TRUE; t1_up := FALSE; 
    ELSIF ((x0 = TRUE) AND  (t0.Q = TRUE) AND  (t1.Q = TRUE)) THEN 
        cstate16 := 42453; y0 := TRUE; y1 := TRUE; y2 := TRUE; t0_start := FALSE;t1_start := TRUE; t1_up := FALSE; 
    END_IF;
17523:
    IF ((x0 = FALSE) AND  (t0.Q = FALSE) AND  (t1.Q = FALSE)) THEN 
        cstate16 := 32883; y0 := FALSE; y1 := FALSE; y2 := FALSE; t0_start := FALSE;t1_start := FALSE; 
    ELSIF ((x0 = FALSE) AND  (t0.Q = FALSE) AND  (t1.Q = TRUE)) THEN 
        cstate16 := 34932; y0 := FALSE; y1 := FALSE; y2 := FALSE; t0_start := FALSE;t1_start := FALSE; 
    ELSIF ((x0 = FALSE) AND  (t0.Q = TRUE) AND  (t1.Q = FALSE)) THEN 
        cstate16 := 27763; y0 := FALSE; y1 := FALSE; y2 := FALSE; t0_start := FALSE;t1_start := FALSE; 
    ELSIF ((x0 = FALSE) AND  (t0.Q = TRUE) AND  (t1.Q = TRUE)) THEN 
        cstate16 := 28788; y0 := FALSE; y1 := FALSE; y2 := FALSE; t0_start := FALSE;t1_start := FALSE; 
    ELSIF ((x0 = TRUE) AND  (t0.Q = FALSE) AND  (t1.Q = FALSE)) THEN 
        cstate16 := 41187; y0 := TRUE; y1 := FALSE; y2 := FALSE; t0_start := TRUE; t0_up := FALSE;t1_start := FALSE; 
    ELSIF ((x0 = TRUE) AND  (t0.Q = FALSE) AND  (t1.Q = TRUE)) THEN 
        cstate16 := 40167; y0 := TRUE; y1 := FALSE; y2 := TRUE; t0_start := TRUE; t0_up := FALSE;t1_start := FALSE; 
    ELSIF ((x0 = TRUE) AND  (t0.Q = TRUE) AND  (t1.Q = FALSE)) THEN 
        cstate16 := 38115; y0 := TRUE; y1 := FALSE; y2 := FALSE; t0_start := TRUE; t0_up := FALSE;t1_start := FALSE; 
    ELSIF ((x0 = TRUE) AND  (t0.Q = TRUE) AND  (t1.Q = TRUE)) THEN 
        cstate16 := 39143; y0 := TRUE; y1 := FALSE; y2 := TRUE; t0_start := TRUE; t0_up := FALSE;t1_start := FALSE; 
    END_IF;
49649:
    IF ((x0 = FALSE) AND  (t0.Q = FALSE) AND  (t1.Q = FALSE)) THEN 
        cstate16 := 32883; y0 := FALSE; y1 := FALSE; y2 := FALSE; t0_start := FALSE;t1_start := FALSE; 
    ELSIF ((x0 = FALSE) AND  (t0.Q = FALSE) AND  (t1.Q = TRUE)) THEN 
        cstate16 := 34932; y0 := FALSE; y1 := FALSE; y2 := FALSE; t0_start := FALSE;t1_start := FALSE; 
    ELSIF ((x0 = FALSE) AND  (t0.Q = TRUE) AND  (t1.Q = FALSE)) THEN 
        cstate16 := 27731; y0 := FALSE; y1 := FALSE; y2 := FALSE; t0_start := FALSE;t1_start := TRUE; t1_up := FALSE; 
    ELSIF ((x0 = FALSE) AND  (t0.Q = TRUE) AND  (t1.Q = TRUE)) THEN 
        cstate16 := 27732; y0 := FALSE; y1 := FALSE; y2 := FALSE; t0_start := FALSE;t1_start := TRUE; t1_up := FALSE; 
    ELSIF ((x0 = TRUE) AND  (t0.Q = FALSE) AND  (t1.Q = FALSE)) THEN 
        cstate16 := 49649; y0 := TRUE; y1 := TRUE; y2 := FALSE; t0_start := FALSE;t1_start := FALSE; 
    ELSIF ((x0 = TRUE) AND  (t0.Q = FALSE) AND  (t1.Q = TRUE)) THEN 
        cstate16 := 48646; y0 := TRUE; y1 := TRUE; y2 := TRUE; t0_start := FALSE;t1_start := FALSE; 
    ELSIF ((x0 = TRUE) AND  (t0.Q = TRUE) AND  (t1.Q = FALSE)) THEN 
        cstate16 := 42449; y0 := TRUE; y1 := TRUE; y2 := FALSE; t0_start := FALSE;t1_start := TRUE; t1_up := FALSE; 
    ELSIF ((x0 = TRUE) AND  (t0.Q = TRUE) AND  (t1.Q = TRUE)) THEN 
        cstate16 := 42453; y0 := TRUE; y1 := TRUE; y2 := TRUE; t0_start := FALSE;t1_start := TRUE; t1_up := FALSE; 
    END_IF;
26130:
    IF ((x0 = FALSE) AND  (t0.Q = FALSE) AND  (t1.Q = FALSE)) THEN 
        cstate16 := 26739; y0 := FALSE; y1 := FALSE; y2 := FALSE; t0_start := FALSE;t1_start := FALSE; 
    ELSIF ((x0 = FALSE) AND  (t0.Q = FALSE) AND  (t1.Q = TRUE)) THEN 
        cstate16 := 26740; y0 := FALSE; y1 := FALSE; y2 := FALSE; t0_start := FALSE;t1_start := FALSE; 
    ELSIF ((x0 = FALSE) AND  (t0.Q = TRUE) AND  (t1.Q = FALSE)) THEN 
        cstate16 := 17491; y0 := FALSE; y1 := FALSE; y2 := FALSE; t0_start := FALSE;t1_start := TRUE; t1_up := FALSE; 
    ELSIF ((x0 = FALSE) AND  (t0.Q = TRUE) AND  (t1.Q = TRUE)) THEN 
        cstate16 := 17492; y0 := FALSE; y1 := FALSE; y2 := FALSE; t0_start := FALSE;t1_start := TRUE; t1_up := FALSE; 
    ELSIF ((x0 = TRUE) AND  (t0.Q = FALSE) AND  (t1.Q = FALSE)) THEN 
        cstate16 := 26129; y0 := TRUE; y1 := TRUE; y2 := FALSE; t0_start := FALSE;t1_start := FALSE; 
    ELSIF ((x0 = TRUE) AND  (t0.Q = FALSE) AND  (t1.Q = TRUE)) THEN 
        cstate16 := 26130; y0 := TRUE; y1 := TRUE; y2 := FALSE; t0_start := FALSE;t1_start := FALSE; 
    ELSIF ((x0 = TRUE) AND  (t0.Q = TRUE) AND  (t1.Q = FALSE)) THEN 
        cstate16 := 42449; y0 := TRUE; y1 := TRUE; y2 := FALSE; t0_start := FALSE;t1_start := TRUE; t1_up := FALSE; 
    ELSIF ((x0 = TRUE) AND  (t0.Q = TRUE) AND  (t1.Q = TRUE)) THEN 
        cstate16 := 42450; y0 := TRUE; y1 := TRUE; y2 := FALSE; t0_start := FALSE;t1_start := TRUE; t1_up := FALSE; 
    END_IF;
48650:
    IF ((x0 = FALSE) AND  (t0.Q = FALSE) AND  (t1.Q = FALSE)) THEN 
        cstate16 := 34931; y0 := FALSE; y1 := FALSE; y2 := FALSE; t0_start := FALSE;t1_start := FALSE; 
    ELSIF ((x0 = FALSE) AND  (t0.Q = FALSE) AND  (t1.Q = TRUE)) THEN 
        cstate16 := 34932; y0 := FALSE; y1 := FALSE; y2 := FALSE; t0_start := FALSE;t1_start := FALSE; 
    ELSIF ((x0 = FALSE) AND  (t0.Q = TRUE) AND  (t1.Q = FALSE)) THEN 
        cstate16 := 27731; y0 := FALSE; y1 := FALSE; y2 := FALSE; t0_start := FALSE;t1_start := TRUE; t1_up := FALSE; 
    ELSIF ((x0 = FALSE) AND  (t0.Q = TRUE) AND  (t1.Q = TRUE)) THEN 
        cstate16 := 27732; y0 := FALSE; y1 := FALSE; y2 := FALSE; t0_start := FALSE;t1_start := TRUE; t1_up := FALSE; 
    ELSIF ((x0 = TRUE) AND  (t0.Q = FALSE) AND  (t1.Q = FALSE)) THEN 
        cstate16 := 48650; y0 := TRUE; y1 := TRUE; y2 := TRUE; t0_start := FALSE;t1_start := FALSE; 
    ELSIF ((x0 = TRUE) AND  (t0.Q = FALSE) AND  (t1.Q = TRUE)) THEN 
        cstate16 := 48646; y0 := TRUE; y1 := TRUE; y2 := TRUE; t0_start := FALSE;t1_start := FALSE; 
    ELSIF ((x0 = TRUE) AND  (t0.Q = TRUE) AND  (t1.Q = FALSE)) THEN 
        cstate16 := 42457; y0 := TRUE; y1 := TRUE; y2 := TRUE; t0_start := FALSE;t1_start := TRUE; t1_up := FALSE; 
    ELSIF ((x0 = TRUE) AND  (t0.Q = TRUE) AND  (t1.Q = TRUE)) THEN 
        cstate16 := 42453; y0 := TRUE; y1 := TRUE; y2 := TRUE; t0_start := FALSE;t1_start := TRUE; t1_up := FALSE; 
    END_IF;
26134:
    IF ((x0 = FALSE) AND  (t0.Q = FALSE) AND  (t1.Q = FALSE)) THEN 
        cstate16 := 26739; y0 := FALSE; y1 := FALSE; y2 := FALSE; t0_start := FALSE;t1_start := FALSE; 
    ELSIF ((x0 = FALSE) AND  (t0.Q = FALSE) AND  (t1.Q = TRUE)) THEN 
        cstate16 := 26740; y0 := FALSE; y1 := FALSE; y2 := FALSE; t0_start := FALSE;t1_start := FALSE; 
    ELSIF ((x0 = FALSE) AND  (t0.Q = TRUE) AND  (t1.Q = FALSE)) THEN 
        cstate16 := 17491; y0 := FALSE; y1 := FALSE; y2 := FALSE; t0_start := FALSE;t1_start := TRUE; t1_up := FALSE; 
    ELSIF ((x0 = FALSE) AND  (t0.Q = TRUE) AND  (t1.Q = TRUE)) THEN 
        cstate16 := 17492; y0 := FALSE; y1 := FALSE; y2 := FALSE; t0_start := FALSE;t1_start := TRUE; t1_up := FALSE; 
    ELSIF ((x0 = TRUE) AND  (t0.Q = FALSE) AND  (t1.Q = FALSE)) THEN 
        cstate16 := 26138; y0 := TRUE; y1 := TRUE; y2 := TRUE; t0_start := FALSE;t1_start := FALSE; 
    ELSIF ((x0 = TRUE) AND  (t0.Q = FALSE) AND  (t1.Q = TRUE)) THEN 
        cstate16 := 26134; y0 := TRUE; y1 := TRUE; y2 := TRUE; t0_start := FALSE;t1_start := FALSE; 
    ELSIF ((x0 = TRUE) AND  (t0.Q = TRUE) AND  (t1.Q = FALSE)) THEN 
        cstate16 := 42457; y0 := TRUE; y1 := TRUE; y2 := TRUE; t0_start := FALSE;t1_start := TRUE; t1_up := FALSE; 
    ELSIF ((x0 = TRUE) AND  (t0.Q = TRUE) AND  (t1.Q = TRUE)) THEN 
        cstate16 := 42453; y0 := TRUE; y1 := TRUE; y2 := TRUE; t0_start := FALSE;t1_start := TRUE; t1_up := FALSE; 
    END_IF;
27732:
    IF ((x0 = FALSE) AND  (t0.Q = FALSE) AND  (t1.Q = FALSE)) THEN 
        cstate16 := 32883; y0 := FALSE; y1 := FALSE; y2 := FALSE; t0_start := FALSE;t1_start := FALSE; 
    ELSIF ((x0 = FALSE) AND  (t0.Q = FALSE) AND  (t1.Q = TRUE)) THEN 
        cstate16 := 34932; y0 := FALSE; y1 := FALSE; y2 := FALSE; t0_start := FALSE;t1_start := FALSE; 
    ELSIF ((x0 = FALSE) AND  (t0.Q = TRUE) AND  (t1.Q = FALSE)) THEN 
        cstate16 := 27763; y0 := FALSE; y1 := FALSE; y2 := FALSE; t0_start := FALSE;t1_start := FALSE; 
    ELSIF ((x0 = FALSE) AND  (t0.Q = TRUE) AND  (t1.Q = TRUE)) THEN 
        cstate16 := 28788; y0 := FALSE; y1 := FALSE; y2 := FALSE; t0_start := FALSE;t1_start := FALSE; 
    ELSIF ((x0 = TRUE) AND  (t0.Q = FALSE) AND  (t1.Q = FALSE)) THEN 
        cstate16 := 41187; y0 := TRUE; y1 := FALSE; y2 := FALSE; t0_start := TRUE; t0_up := FALSE;t1_start := FALSE; 
    ELSIF ((x0 = TRUE) AND  (t0.Q = FALSE) AND  (t1.Q = TRUE)) THEN 
        cstate16 := 40164; y0 := TRUE; y1 := FALSE; y2 := FALSE; t0_start := TRUE; t0_up := FALSE;t1_start := FALSE; 
